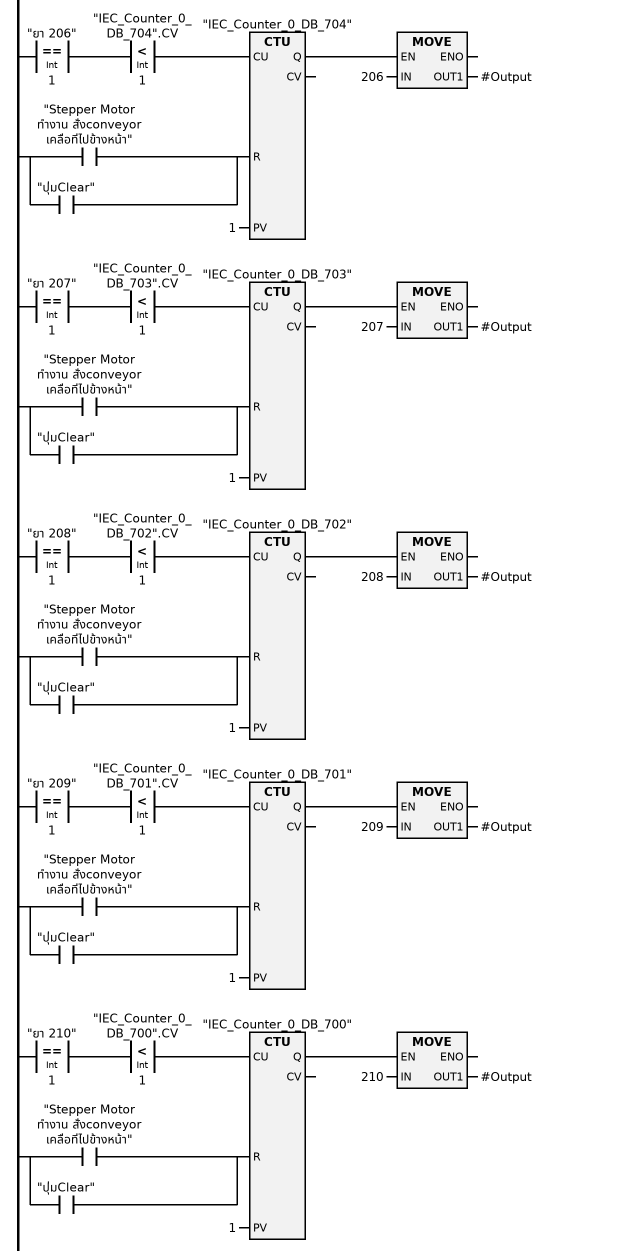
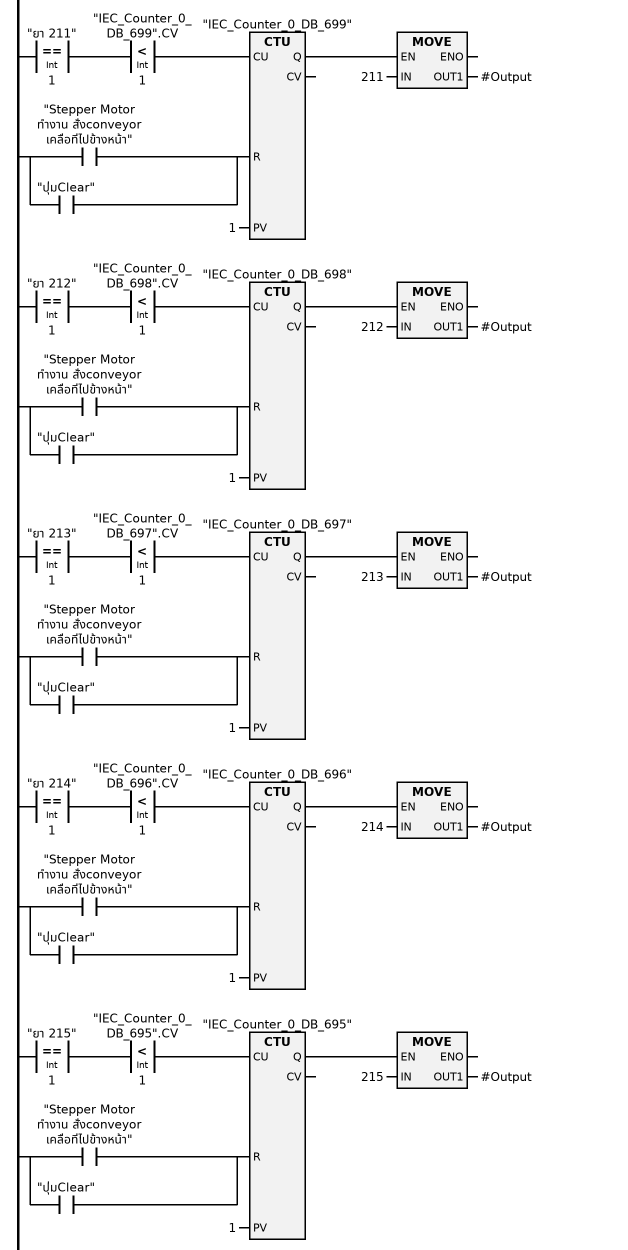
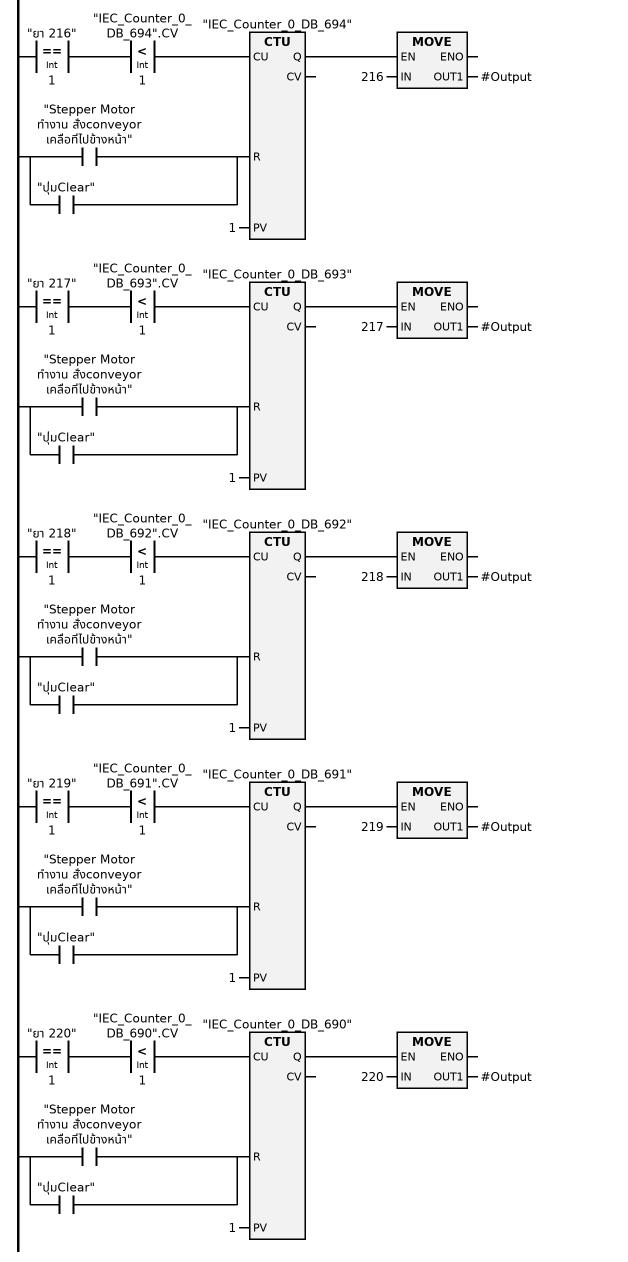
   "IEC_Counter_0_DB_709".CTU(CU := ("ยา 201" = 1) AND ("IEC_Counter_0_DB_709".CV < 1),
                           R := "Stepper Motor ทำงาน สั่งconveyor เคลื่อที่ไปข้างหน้า" OR "ปุ่มClear",
                           PV := 1);
   IF "IEC_Counter_0_DB_709".Q THEN #Output := 201; END_IF;
   "IEC_Counter_0_DB_705".CTU(CU := ("ยา 202" = 1) AND ("IEC_Counter_0_DB_705".CV < 1),
                           R := "Stepper Motor ทำงาน สั่งconveyor เคลื่อที่ไปข้างหน้า" OR "ปุ่มClear",
                           PV := 1);
   IF "IEC_Counter_0_DB_705".Q THEN #Output := 202; END_IF;
   "IEC_Counter_0_DB_708".CTU(CU := ("ยา 203" = 1) AND ("IEC_Counter_0_DB_708".CV < 1),
                           R := "Stepper Motor ทำงาน สั่งconveyor เคลื่อที่ไปข้างหน้า" OR "ปุ่มClear",
                           PV := 1);
   IF "IEC_Counter_0_DB_708".Q THEN #Output := 203; END_IF;
   "IEC_Counter_0_DB_707".CTU(CU := ("ยา 204" = 1) AND ("IEC_Counter_0_DB_707".CV < 1),
                           R := "Stepper Motor ทำงาน สั่งconveyor เคลื่อที่ไปข้างหน้า" OR "ปุ่มClear",
                           PV := 1);
   IF "IEC_Counter_0_DB_707".Q THEN #Output := 204; END_IF;
   "IEC_Counter_0_DB_706".CTU(CU := ("ยา 205" = 1) AND ("IEC_Counter_0_DB_706".CV < 1),
                           R := "Stepper Motor ทำงาน สั่งconveyor เคลื่อที่ไปข้างหน้า" OR "ปุ่มClear",
                           PV := 1);
   IF "IEC_Counter_0_DB_706".Q THEN #Output := 205; END_IF;
   "IEC_Counter_0_DB_704".CTU(CU := ("ยา 206" = 1) AND ("IEC_Counter_0_DB_704".CV < 1),
                           R := "Stepper Motor ทำงาน สั่งconveyor เคลื่อที่ไปข้างหน้า" OR "ปุ่มClear",
                           PV := 1);
   IF "IEC_Counter_0_DB_704".Q THEN #Output := 206; END_IF;
   "IEC_Counter_0_DB_703".CTU(CU := ("ยา 207" = 1) AND ("IEC_Counter_0_DB_703".CV < 1),
                           R := "Stepper Motor ทำงาน สั่งconveyor เคลื่อที่ไปข้างหน้า" OR "ปุ่มClear",
                           PV := 1);
   IF "IEC_Counter_0_DB_703".Q THEN #Output := 207; END_IF;
   "IEC_Counter_0_DB_702".CTU(CU := ("ยา 208" = 1) AND ("IEC_Counter_0_DB_702".CV < 1),
                           R := "Stepper Motor ทำงาน สั่งconveyor เคลื่อที่ไปข้างหน้า" OR "ปุ่มClear",
                           PV := 1);
   IF "IEC_Counter_0_DB_702".Q THEN #Output := 208; END_IF;
   "IEC_Counter_0_DB_701".CTU(CU := ("ยา 209" = 1) AND ("IEC_Counter_0_DB_701".CV < 1),
                           R := "Stepper Motor ทำงาน สั่งconveyor เคลื่อที่ไปข้างหน้า" OR "ปุ่มClear",
                           PV := 1);
   IF "IEC_Counter_0_DB_701".Q THEN #Output := 209; END_IF;
   "IEC_Counter_0_DB_700".CTU(CU := ("ยา 210" = 1) AND ("IEC_Counter_0_DB_700".CV < 1),
                           R := "Stepper Motor ทำงาน สั่งconveyor เคลื่อที่ไปข้างหน้า" OR "ปุ่มClear",
                           PV := 1);
   IF "IEC_Counter_0_DB_700".Q THEN #Output := 210; END_IF;
   "IEC_Counter_0_DB_699".CTU(CU := ("ยา 211" = 1) AND ("IEC_Counter_0_DB_699".CV < 1),
                           R := "Stepper Motor ทำงาน สั่งconveyor เคลื่อที่ไปข้างหน้า" OR "ปุ่มClear",
                           PV := 1);
   IF "IEC_Counter_0_DB_699".Q THEN #Output := 211; END_IF;
   "IEC_Counter_0_DB_698".CTU(CU := ("ยา 212" = 1) AND ("IEC_Counter_0_DB_698".CV < 1),
                           R := "Stepper Motor ทำงาน สั่งconveyor เคลื่อที่ไปข้างหน้า" OR "ปุ่มClear",
                           PV := 1);
   IF "IEC_Counter_0_DB_698".Q THEN #Output := 212; END_IF;
   "IEC_Counter_0_DB_697".CTU(CU := ("ยา 213" = 1) AND ("IEC_Counter_0_DB_697".CV < 1),
                           R := "Stepper Motor ทำงาน สั่งconveyor เคลื่อที่ไปข้างหน้า" OR "ปุ่มClear",
                           PV := 1);
   IF "IEC_Counter_0_DB_697".Q THEN #Output := 213; END_IF;
   "IEC_Counter_0_DB_696".CTU(CU := ("ยา 214" = 1) AND ("IEC_Counter_0_DB_696".CV < 1),
                           R := "Stepper Motor ทำงาน สั่งconveyor เคลื่อที่ไปข้างหน้า" OR "ปุ่มClear",
                           PV := 1);
   IF "IEC_Counter_0_DB_696".Q THEN #Output := 214; END_IF;
   "IEC_Counter_0_DB_695".CTU(CU := ("ยา 215" = 1) AND ("IEC_Counter_0_DB_695".CV < 1),
                           R := "Stepper Motor ทำงาน สั่งconveyor เคลื่อที่ไปข้างหน้า" OR "ปุ่มClear",
                           PV := 1);
   IF "IEC_Counter_0_DB_695".Q THEN #Output := 215; END_IF;
   "IEC_Counter_0_DB_694".CTU(CU := ("ยา 216" = 1) AND ("IEC_Counter_0_DB_694".CV < 1),
                           R := "Stepper Motor ทำงาน สั่งconveyor เคลื่อที่ไปข้างหน้า" OR "ปุ่มClear",
                           PV := 1);
   IF "IEC_Counter_0_DB_694".Q THEN #Output := 216; END_IF;
   "IEC_Counter_0_DB_693".CTU(CU := ("ยา 217" = 1) AND ("IEC_Counter_0_DB_693".CV < 1),
                           R := "Stepper Motor ทำงาน สั่งconveyor เคลื่อที่ไปข้างหน้า" OR "ปุ่มClear",
                           PV := 1);
   IF "IEC_Counter_0_DB_693".Q THEN #Output := 217; END_IF;
   "IEC_Counter_0_DB_692".CTU(CU := ("ยา 218" = 1) AND ("IEC_Counter_0_DB_692".CV < 1),
                           R := "Stepper Motor ทำงาน สั่งconveyor เคลื่อที่ไปข้างหน้า" OR "ปุ่มClear",
                           PV := 1);
   IF "IEC_Counter_0_DB_692".Q THEN #Output := 218; END_IF;
   "IEC_Counter_0_DB_691".CTU(CU := ("ยา 219" = 1) AND ("IEC_Counter_0_DB_691".CV < 1),
                           R := "Stepper Motor ทำงาน สั่งconveyor เคลื่อที่ไปข้างหน้า" OR "ปุ่มClear",
                           PV := 1);
   IF "IEC_Counter_0_DB_691".Q THEN #Output := 219; END_IF;
   "IEC_Counter_0_DB_690".CTU(CU := ("ยา 220" = 1) AND ("IEC_Counter_0_DB_690".CV < 1),
                           R := "Stepper Motor ทำงาน สั่งconveyor เคลื่อที่ไปข้างหน้า" OR "ปุ่มClear",
                           PV := 1);
   IF "IEC_Counter_0_DB_690".Q THEN #Output := 220; END_IF;
END_REGION

REGION Network 12
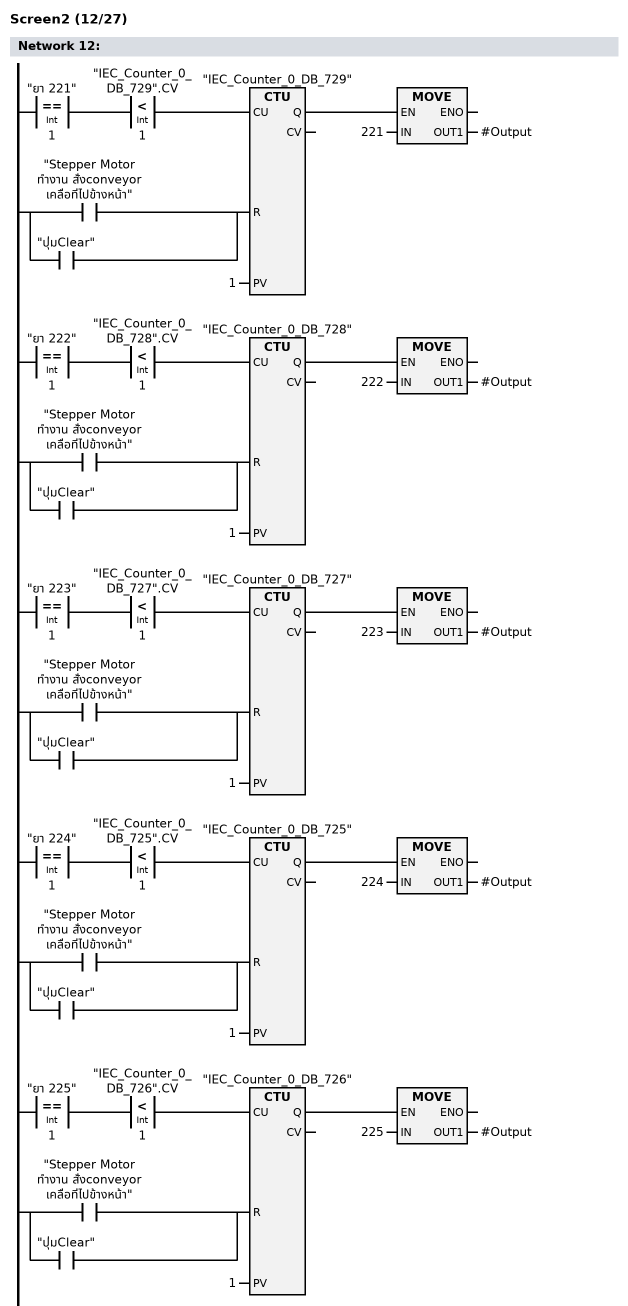
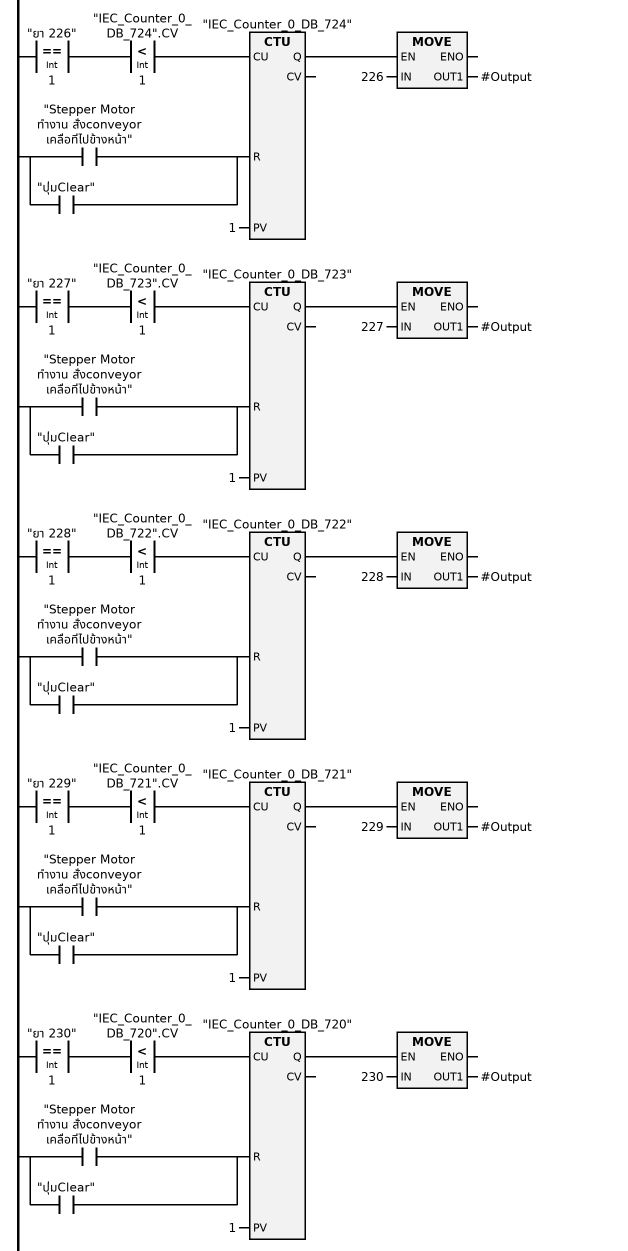
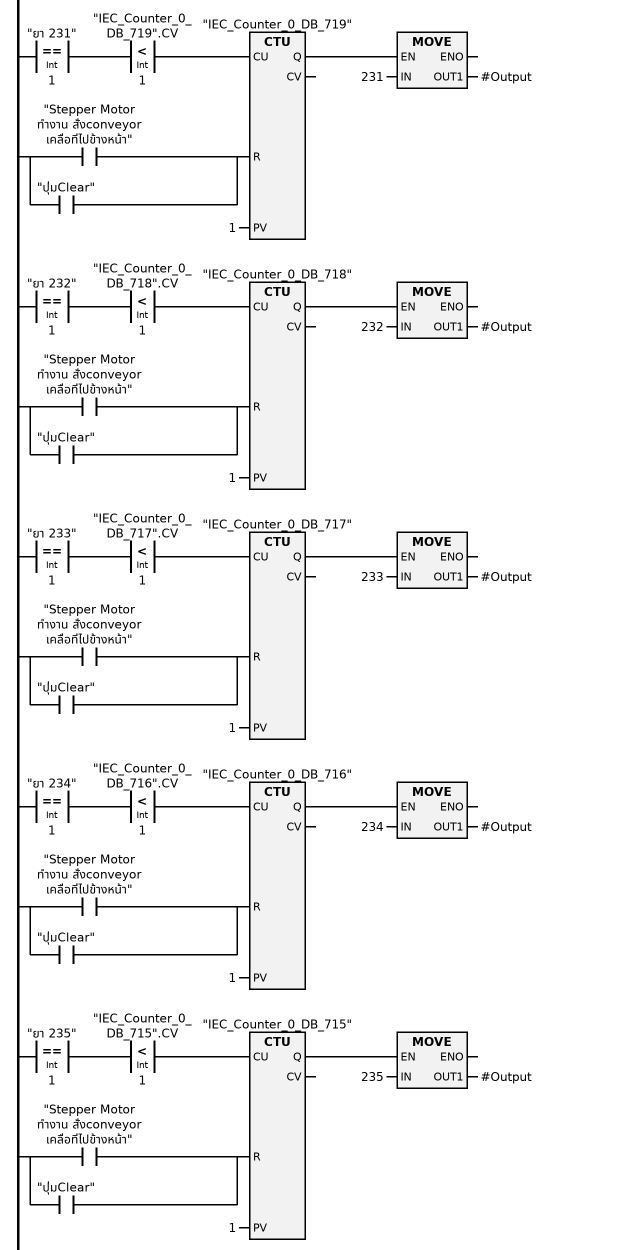
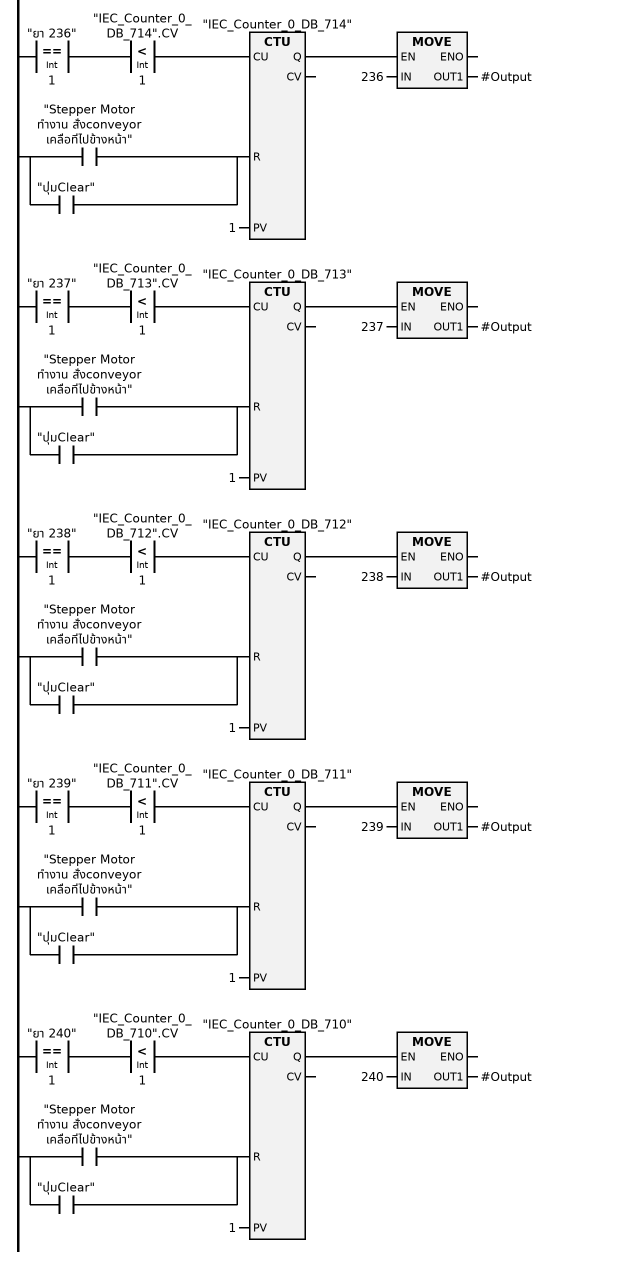
   "IEC_Counter_0_DB_729".CTU(CU := ("ยา 221" = 1) AND ("IEC_Counter_0_DB_729".CV < 1),
                           R := "Stepper Motor ทำงาน สั่งconveyor เคลื่อที่ไปข้างหน้า" OR "ปุ่มClear",
                           PV := 1);
   IF "IEC_Counter_0_DB_729".Q THEN #Output := 221; END_IF;
   "IEC_Counter_0_DB_728".CTU(CU := ("ยา 222" = 1) AND ("IEC_Counter_0_DB_728".CV < 1),
                           R := "Stepper Motor ทำงาน สั่งconveyor เคลื่อที่ไปข้างหน้า" OR "ปุ่มClear",
                           PV := 1);
   IF "IEC_Counter_0_DB_728".Q THEN #Output := 222; END_IF;
   "IEC_Counter_0_DB_727".CTU(CU := ("ยา 223" = 1) AND ("IEC_Counter_0_DB_727".CV < 1),
                           R := "Stepper Motor ทำงาน สั่งconveyor เคลื่อที่ไปข้างหน้า" OR "ปุ่มClear",
                           PV := 1);
   IF "IEC_Counter_0_DB_727".Q THEN #Output := 223; END_IF;
   "IEC_Counter_0_DB_725".CTU(CU := ("ยา 224" = 1) AND ("IEC_Counter_0_DB_725".CV < 1),
                           R := "Stepper Motor ทำงาน สั่งconveyor เคลื่อที่ไปข้างหน้า" OR "ปุ่มClear",
                           PV := 1);
   IF "IEC_Counter_0_DB_725".Q THEN #Output := 224; END_IF;
   "IEC_Counter_0_DB_726".CTU(CU := ("ยา 225" = 1) AND ("IEC_Counter_0_DB_726".CV < 1),
                           R := "Stepper Motor ทำงาน สั่งconveyor เคลื่อที่ไปข้างหน้า" OR "ปุ่มClear",
                           PV := 1);
   IF "IEC_Counter_0_DB_726".Q THEN #Output := 225; END_IF;
   "IEC_Counter_0_DB_724".CTU(CU := ("ยา 226" = 1) AND ("IEC_Counter_0_DB_724".CV < 1),
                           R := "Stepper Motor ทำงาน สั่งconveyor เคลื่อที่ไปข้างหน้า" OR "ปุ่มClear",
                           PV := 1);
   IF "IEC_Counter_0_DB_724".Q THEN #Output := 226; END_IF;
   "IEC_Counter_0_DB_723".CTU(CU := ("ยา 227" = 1) AND ("IEC_Counter_0_DB_723".CV < 1),
                           R := "Stepper Motor ทำงาน สั่งconveyor เคลื่อที่ไปข้างหน้า" OR "ปุ่มClear",
                           PV := 1);
   IF "IEC_Counter_0_DB_723".Q THEN #Output := 227; END_IF;
   "IEC_Counter_0_DB_722".CTU(CU := ("ยา 228" = 1) AND ("IEC_Counter_0_DB_722".CV < 1),
                           R := "Stepper Motor ทำงาน สั่งconveyor เคลื่อที่ไปข้างหน้า" OR "ปุ่มClear",
                           PV := 1);
   IF "IEC_Counter_0_DB_722".Q THEN #Output := 228; END_IF;
   "IEC_Counter_0_DB_721".CTU(CU := ("ยา 229" = 1) AND ("IEC_Counter_0_DB_721".CV < 1),
                           R := "Stepper Motor ทำงาน สั่งconveyor เคลื่อที่ไปข้างหน้า" OR "ปุ่มClear",
                           PV := 1);
   IF "IEC_Counter_0_DB_721".Q THEN #Output := 229; END_IF;
   "IEC_Counter_0_DB_720".CTU(CU := ("ยา 230" = 1) AND ("IEC_Counter_0_DB_720".CV < 1),
                           R := "Stepper Motor ทำงาน สั่งconveyor เคลื่อที่ไปข้างหน้า" OR "ปุ่มClear",
                           PV := 1);
   IF "IEC_Counter_0_DB_720".Q THEN #Output := 230; END_IF;
   "IEC_Counter_0_DB_719".CTU(CU := ("ยา 231" = 1) AND ("IEC_Counter_0_DB_719".CV < 1),
                           R := "Stepper Motor ทำงาน สั่งconveyor เคลื่อที่ไปข้างหน้า" OR "ปุ่มClear",
                           PV := 1);
   IF "IEC_Counter_0_DB_719".Q THEN #Output := 231; END_IF;
   "IEC_Counter_0_DB_718".CTU(CU := ("ยา 232" = 1) AND ("IEC_Counter_0_DB_718".CV < 1),
                           R := "Stepper Motor ทำงาน สั่งconveyor เคลื่อที่ไปข้างหน้า" OR "ปุ่มClear",
                           PV := 1);
   IF "IEC_Counter_0_DB_718".Q THEN #Output := 232; END_IF;
   "IEC_Counter_0_DB_717".CTU(CU := ("ยา 233" = 1) AND ("IEC_Counter_0_DB_717".CV < 1),
                           R := "Stepper Motor ทำงาน สั่งconveyor เคลื่อที่ไปข้างหน้า" OR "ปุ่มClear",
                           PV := 1);
   IF "IEC_Counter_0_DB_717".Q THEN #Output := 233; END_IF;
   "IEC_Counter_0_DB_716".CTU(CU := ("ยา 234" = 1) AND ("IEC_Counter_0_DB_716".CV < 1),
                           R := "Stepper Motor ทำงาน สั่งconveyor เคลื่อที่ไปข้างหน้า" OR "ปุ่มClear",
                           PV := 1);
   IF "IEC_Counter_0_DB_716".Q THEN #Output := 234; END_IF;
   "IEC_Counter_0_DB_715".CTU(CU := ("ยา 235" = 1) AND ("IEC_Counter_0_DB_715".CV < 1),
                           R := "Stepper Motor ทำงาน สั่งconveyor เคลื่อที่ไปข้างหน้า" OR "ปุ่มClear",
                           PV := 1);
   IF "IEC_Counter_0_DB_715".Q THEN #Output := 235; END_IF;
   "IEC_Counter_0_DB_714".CTU(CU := ("ยา 236" = 1) AND ("IEC_Counter_0_DB_714".CV < 1),
                           R := "Stepper Motor ทำงาน สั่งconveyor เคลื่อที่ไปข้างหน้า" OR "ปุ่มClear",
                           PV := 1);
   IF "IEC_Counter_0_DB_714".Q THEN #Output := 236; END_IF;
   "IEC_Counter_0_DB_713".CTU(CU := ("ยา 237" = 1) AND ("IEC_Counter_0_DB_713".CV < 1),
                           R := "Stepper Motor ทำงาน สั่งconveyor เคลื่อที่ไปข้างหน้า" OR "ปุ่มClear",
                           PV := 1);
   IF "IEC_Counter_0_DB_713".Q THEN #Output := 237; END_IF;
   "IEC_Counter_0_DB_712".CTU(CU := ("ยา 238" = 1) AND ("IEC_Counter_0_DB_712".CV < 1),
                           R := "Stepper Motor ทำงาน สั่งconveyor เคลื่อที่ไปข้างหน้า" OR "ปุ่มClear",
                           PV := 1);
   IF "IEC_Counter_0_DB_712".Q THEN #Output := 238; END_IF;
   "IEC_Counter_0_DB_711".CTU(CU := ("ยา 239" = 1) AND ("IEC_Counter_0_DB_711".CV < 1),
                           R := "Stepper Motor ทำงาน สั่งconveyor เคลื่อที่ไปข้างหน้า" OR "ปุ่มClear",
                           PV := 1);
   IF "IEC_Counter_0_DB_711".Q THEN #Output := 239; END_IF;
   "IEC_Counter_0_DB_710".CTU(CU := ("ยา 240" = 1) AND ("IEC_Counter_0_DB_710".CV < 1),
                           R := "Stepper Motor ทำงาน สั่งconveyor เคลื่อที่ไปข้างหน้า" OR "ปุ่มClear",
                           PV := 1);
   IF "IEC_Counter_0_DB_710".Q THEN #Output := 240; END_IF;
END_REGION

REGION Network 13
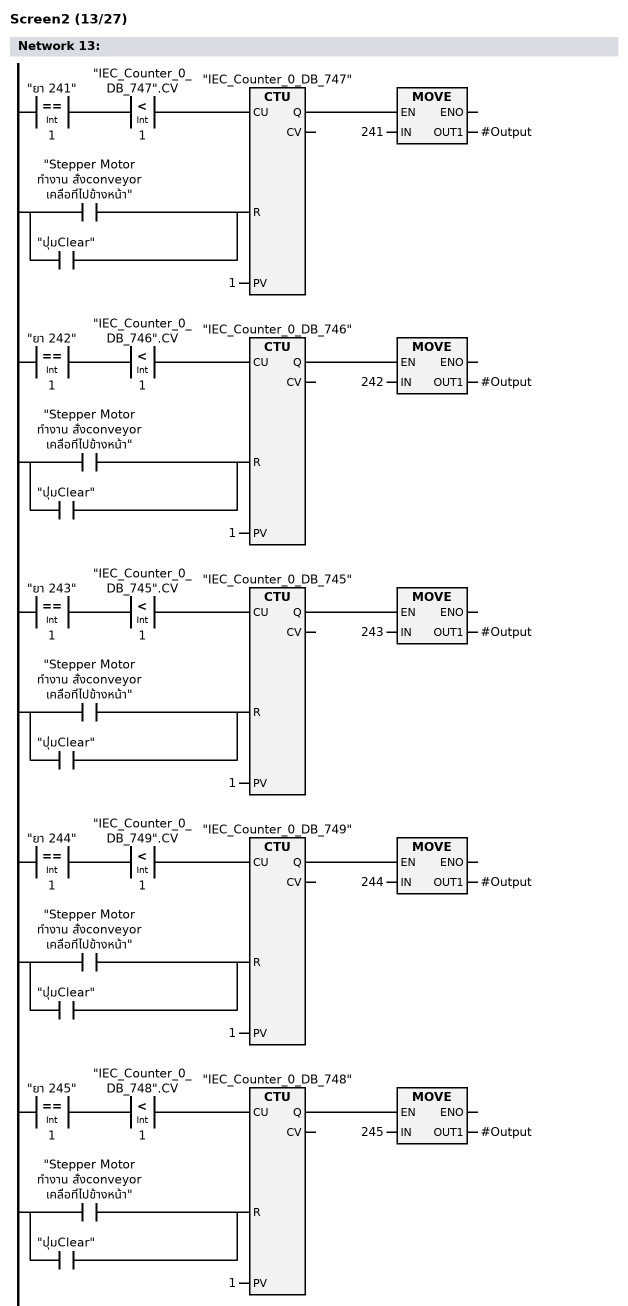
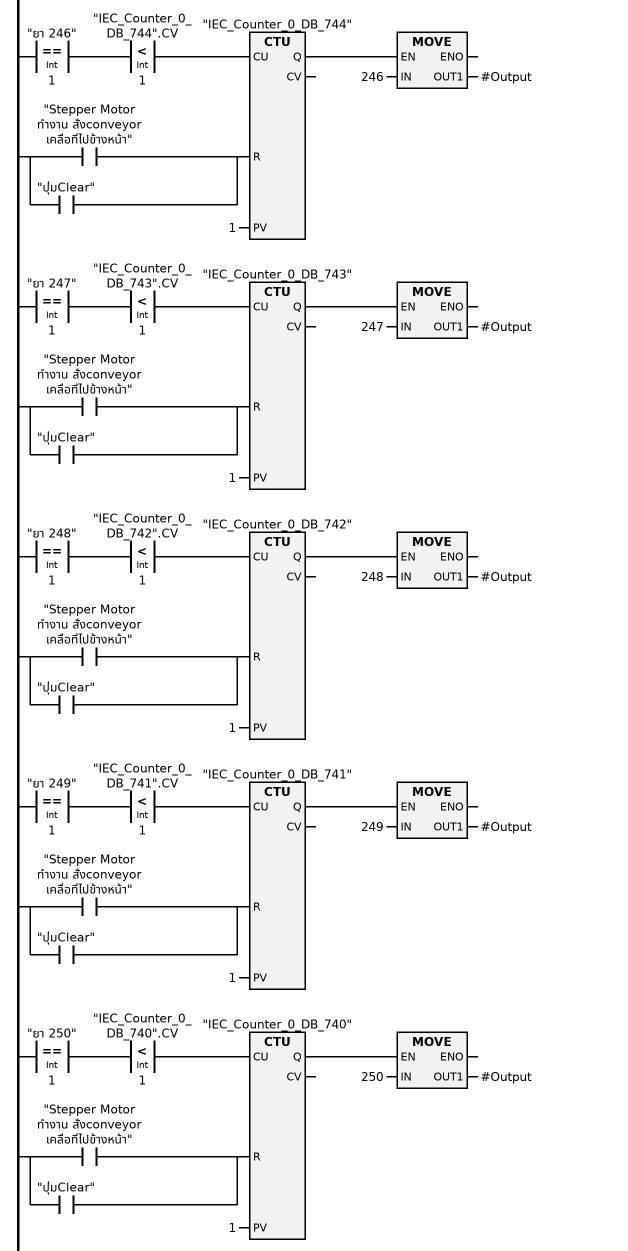
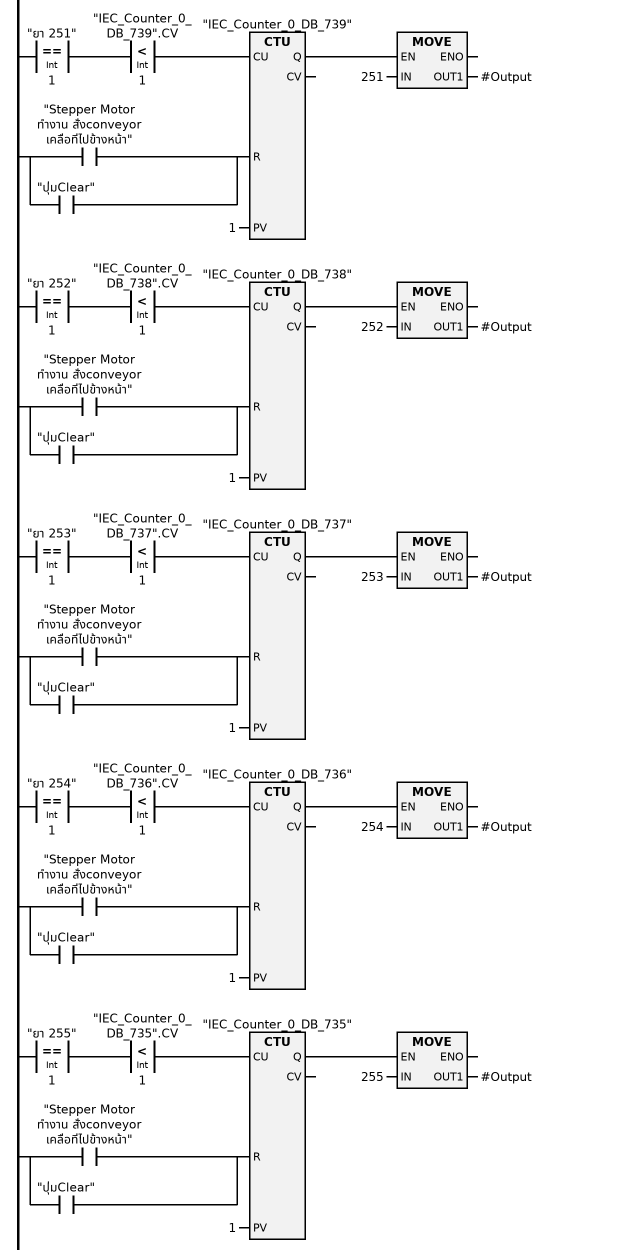
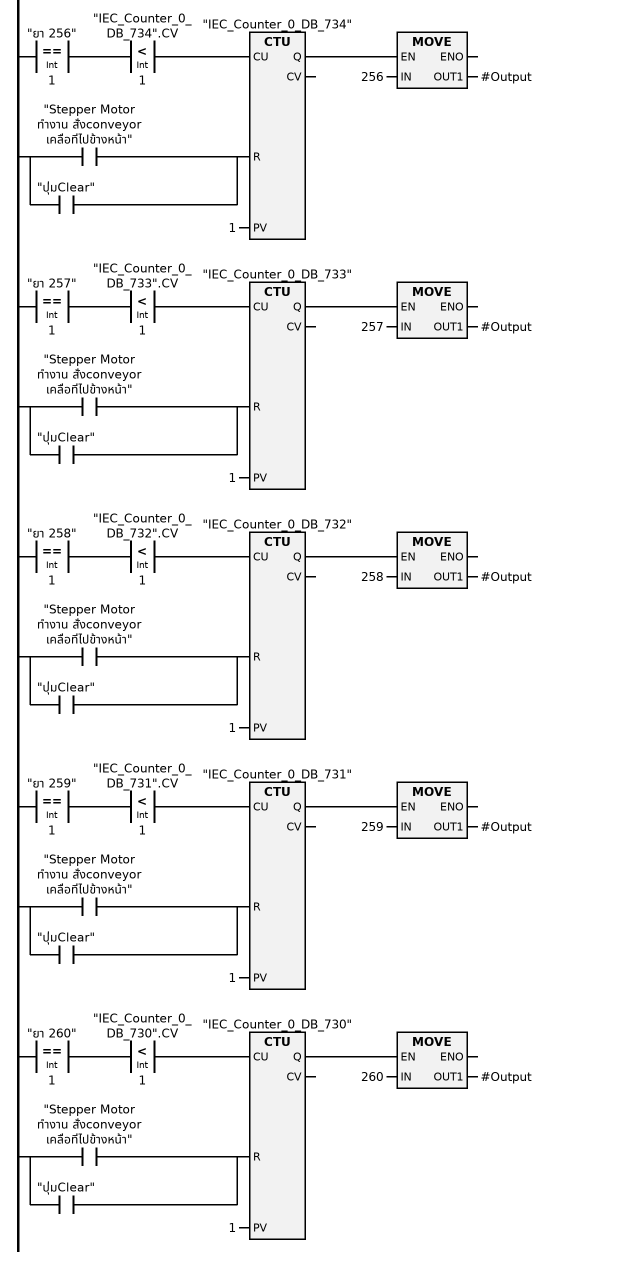
   "IEC_Counter_0_DB_747".CTU(CU := ("ยา 241" = 1) AND ("IEC_Counter_0_DB_747".CV < 1),
                           R := "Stepper Motor ทำงาน สั่งconveyor เคลื่อที่ไปข้างหน้า" OR "ปุ่มClear",
                           PV := 1);
   IF "IEC_Counter_0_DB_747".Q THEN #Output := 241; END_IF;
   "IEC_Counter_0_DB_746".CTU(CU := ("ยา 242" = 1) AND ("IEC_Counter_0_DB_746".CV < 1),
                           R := "Stepper Motor ทำงาน สั่งconveyor เคลื่อที่ไปข้างหน้า" OR "ปุ่มClear",
                           PV := 1);
   IF "IEC_Counter_0_DB_746".Q THEN #Output := 242; END_IF;
   "IEC_Counter_0_DB_745".CTU(CU := ("ยา 243" = 1) AND ("IEC_Counter_0_DB_745".CV < 1),
                           R := "Stepper Motor ทำงาน สั่งconveyor เคลื่อที่ไปข้างหน้า" OR "ปุ่มClear",
                           PV := 1);
   IF "IEC_Counter_0_DB_745".Q THEN #Output := 243; END_IF;
   "IEC_Counter_0_DB_749".CTU(CU := ("ยา 244" = 1) AND ("IEC_Counter_0_DB_749".CV < 1),
                           R := "Stepper Motor ทำงาน สั่งconveyor เคลื่อที่ไปข้างหน้า" OR "ปุ่มClear",
                           PV := 1);
   IF "IEC_Counter_0_DB_749".Q THEN #Output := 244; END_IF;
   "IEC_Counter_0_DB_748".CTU(CU := ("ยา 245" = 1) AND ("IEC_Counter_0_DB_748".CV < 1),
                           R := "Stepper Motor ทำงาน สั่งconveyor เคลื่อที่ไปข้างหน้า" OR "ปุ่มClear",
                           PV := 1);
   IF "IEC_Counter_0_DB_748".Q THEN #Output := 245; END_IF;
   "IEC_Counter_0_DB_744".CTU(CU := ("ยา 246" = 1) AND ("IEC_Counter_0_DB_744".CV < 1),
                           R := "Stepper Motor ทำงาน สั่งconveyor เคลื่อที่ไปข้างหน้า" OR "ปุ่มClear",
                           PV := 1);
   IF "IEC_Counter_0_DB_744".Q THEN #Output := 246; END_IF;
   "IEC_Counter_0_DB_743".CTU(CU := ("ยา 247" = 1) AND ("IEC_Counter_0_DB_743".CV < 1),
                           R := "Stepper Motor ทำงาน สั่งconveyor เคลื่อที่ไปข้างหน้า" OR "ปุ่มClear",
                           PV := 1);
   IF "IEC_Counter_0_DB_743".Q THEN #Output := 247; END_IF;
   "IEC_Counter_0_DB_742".CTU(CU := ("ยา 248" = 1) AND ("IEC_Counter_0_DB_742".CV < 1),
                           R := "Stepper Motor ทำงาน สั่งconveyor เคลื่อที่ไปข้างหน้า" OR "ปุ่มClear",
                           PV := 1);
   IF "IEC_Counter_0_DB_742".Q THEN #Output := 248; END_IF;
   "IEC_Counter_0_DB_741".CTU(CU := ("ยา 249" = 1) AND ("IEC_Counter_0_DB_741".CV < 1),
                           R := "Stepper Motor ทำงาน สั่งconveyor เคลื่อที่ไปข้างหน้า" OR "ปุ่มClear",
                           PV := 1);
   IF "IEC_Counter_0_DB_741".Q THEN #Output := 249; END_IF;
   "IEC_Counter_0_DB_740".CTU(CU := ("ยา 250" = 1) AND ("IEC_Counter_0_DB_740".CV < 1),
                           R := "Stepper Motor ทำงาน สั่งconveyor เคลื่อที่ไปข้างหน้า" OR "ปุ่มClear",
                           PV := 1);
   IF "IEC_Counter_0_DB_740".Q THEN #Output := 250; END_IF;
   "IEC_Counter_0_DB_739".CTU(CU := ("ยา 251" = 1) AND ("IEC_Counter_0_DB_739".CV < 1),
                           R := "Stepper Motor ทำงาน สั่งconveyor เคลื่อที่ไปข้างหน้า" OR "ปุ่มClear",
                           PV := 1);
   IF "IEC_Counter_0_DB_739".Q THEN #Output := 251; END_IF;
   "IEC_Counter_0_DB_738".CTU(CU := ("ยา 252" = 1) AND ("IEC_Counter_0_DB_738".CV < 1),
                           R := "Stepper Motor ทำงาน สั่งconveyor เคลื่อที่ไปข้างหน้า" OR "ปุ่มClear",
                           PV := 1);
   IF "IEC_Counter_0_DB_738".Q THEN #Output := 252; END_IF;
   "IEC_Counter_0_DB_737".CTU(CU := ("ยา 253" = 1) AND ("IEC_Counter_0_DB_737".CV < 1),
                           R := "Stepper Motor ทำงาน สั่งconveyor เคลื่อที่ไปข้างหน้า" OR "ปุ่มClear",
                           PV := 1);
   IF "IEC_Counter_0_DB_737".Q THEN #Output := 253; END_IF;
   "IEC_Counter_0_DB_736".CTU(CU := ("ยา 254" = 1) AND ("IEC_Counter_0_DB_736".CV < 1),
                           R := "Stepper Motor ทำงาน สั่งconveyor เคลื่อที่ไปข้างหน้า" OR "ปุ่มClear",
                           PV := 1);
   IF "IEC_Counter_0_DB_736".Q THEN #Output := 254; END_IF;
   "IEC_Counter_0_DB_735".CTU(CU := ("ยา 255" = 1) AND ("IEC_Counter_0_DB_735".CV < 1),
                           R := "Stepper Motor ทำงาน สั่งconveyor เคลื่อที่ไปข้างหน้า" OR "ปุ่มClear",
                           PV := 1);
   IF "IEC_Counter_0_DB_735".Q THEN #Output := 255; END_IF;
   "IEC_Counter_0_DB_734".CTU(CU := ("ยา 256" = 1) AND ("IEC_Counter_0_DB_734".CV < 1),
                           R := "Stepper Motor ทำงาน สั่งconveyor เคลื่อที่ไปข้างหน้า" OR "ปุ่มClear",
                           PV := 1);
   IF "IEC_Counter_0_DB_734".Q THEN #Output := 256; END_IF;
   "IEC_Counter_0_DB_733".CTU(CU := ("ยา 257" = 1) AND ("IEC_Counter_0_DB_733".CV < 1),
                           R := "Stepper Motor ทำงาน สั่งconveyor เคลื่อที่ไปข้างหน้า" OR "ปุ่มClear",
                           PV := 1);
   IF "IEC_Counter_0_DB_733".Q THEN #Output := 257; END_IF;
   "IEC_Counter_0_DB_732".CTU(CU := ("ยา 258" = 1) AND ("IEC_Counter_0_DB_732".CV < 1),
                           R := "Stepper Motor ทำงาน สั่งconveyor เคลื่อที่ไปข้างหน้า" OR "ปุ่มClear",
                           PV := 1);
   IF "IEC_Counter_0_DB_732".Q THEN #Output := 258; END_IF;
   "IEC_Counter_0_DB_731".CTU(CU := ("ยา 259" = 1) AND ("IEC_Counter_0_DB_731".CV < 1),
                           R := "Stepper Motor ทำงาน สั่งconveyor เคลื่อที่ไปข้างหน้า" OR "ปุ่มClear",
                           PV := 1);
   IF "IEC_Counter_0_DB_731".Q THEN #Output := 259; END_IF;
   "IEC_Counter_0_DB_730".CTU(CU := ("ยา 260" = 1) AND ("IEC_Counter_0_DB_730".CV < 1),
                           R := "Stepper Motor ทำงาน สั่งconveyor เคลื่อที่ไปข้างหน้า" OR "ปุ่มClear",
                           PV := 1);
   IF "IEC_Counter_0_DB_730".Q THEN #Output := 260; END_IF;
END_REGION

REGION Network 14
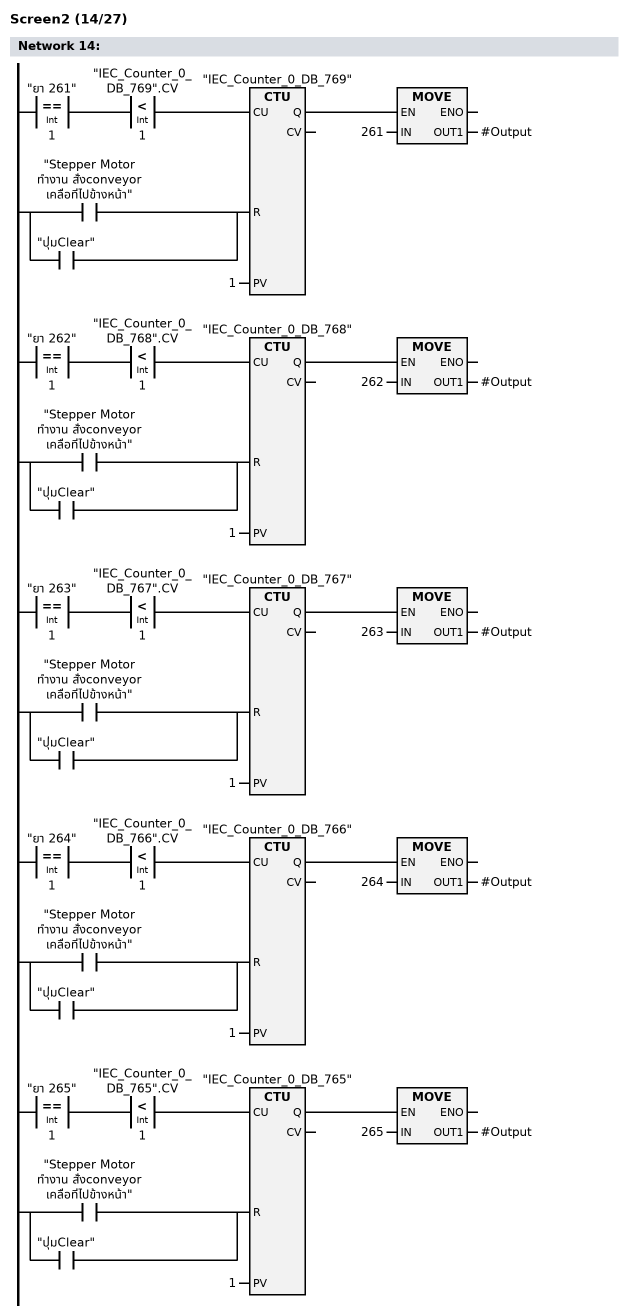
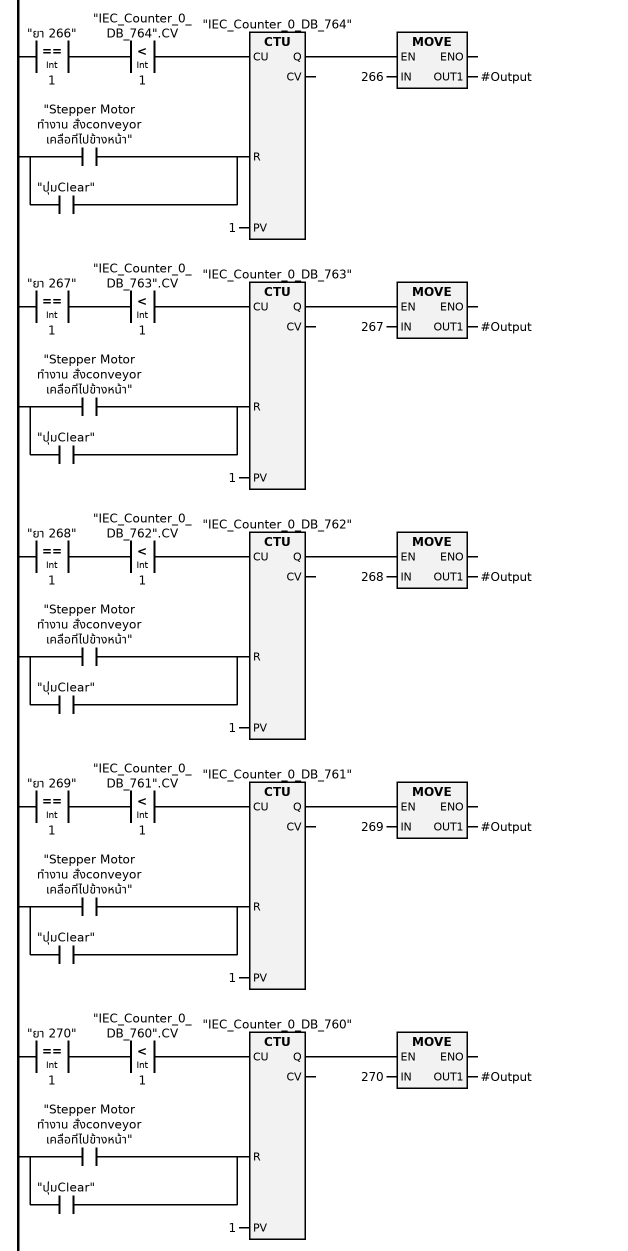
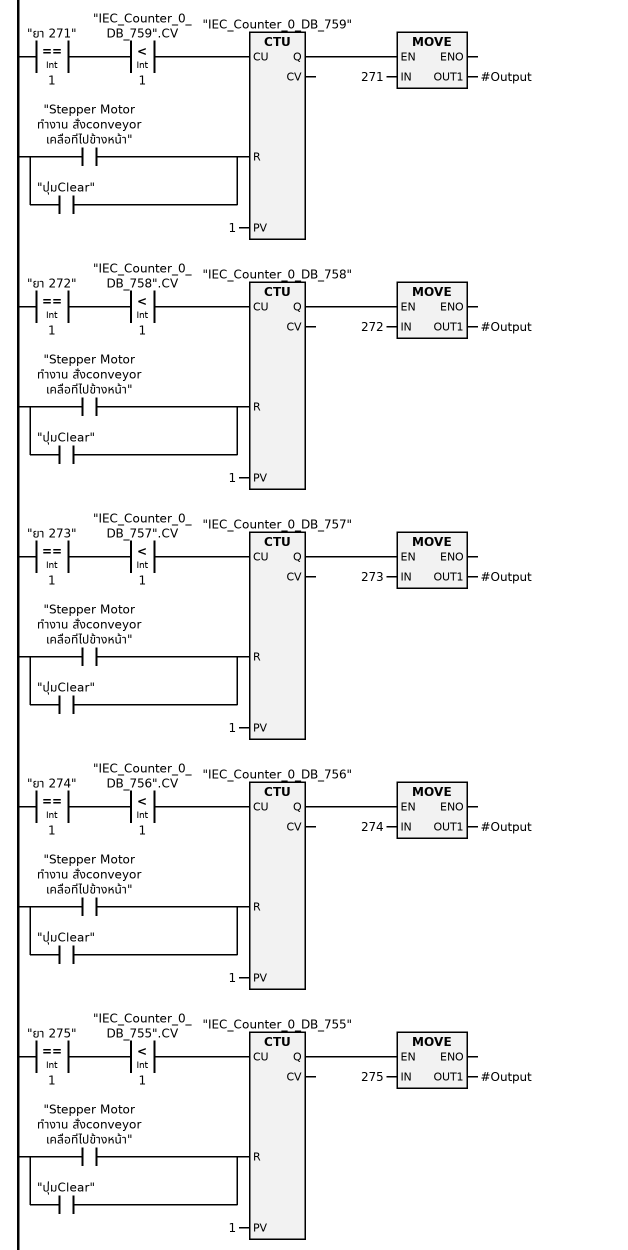
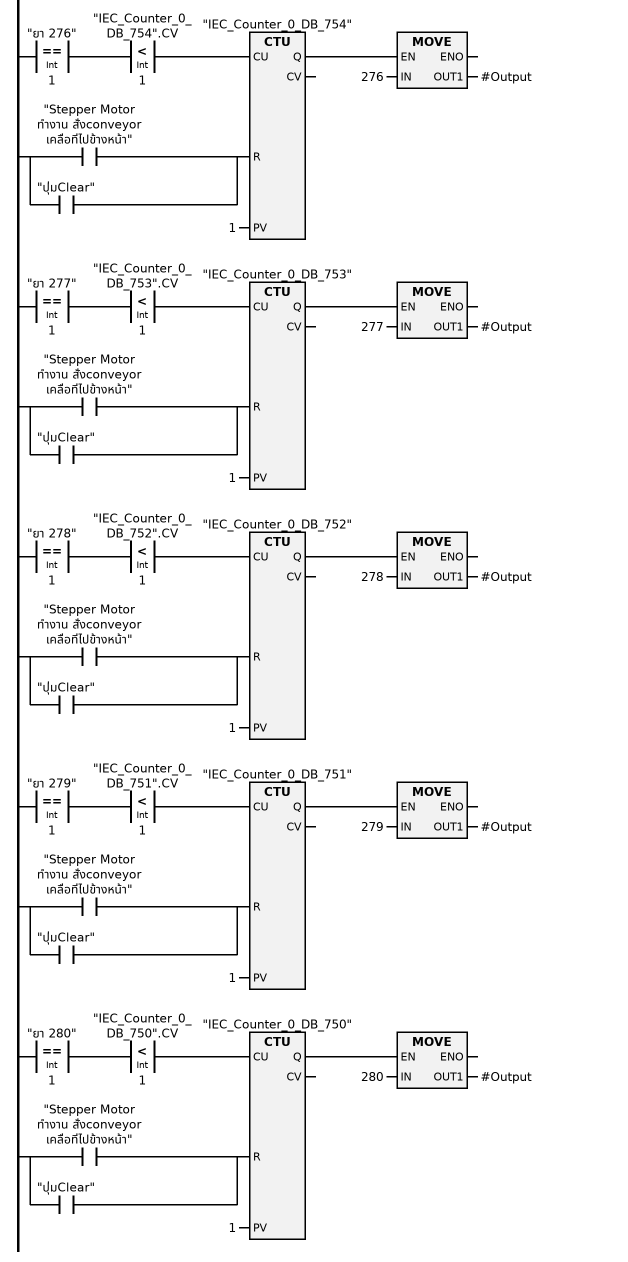
   "IEC_Counter_0_DB_769".CTU(CU := ("ยา 261" = 1) AND ("IEC_Counter_0_DB_769".CV < 1),
                           R := "Stepper Motor ทำงาน สั่งconveyor เคลื่อที่ไปข้างหน้า" OR "ปุ่มClear",
                           PV := 1);
   IF "IEC_Counter_0_DB_769".Q THEN #Output := 261; END_IF;
   "IEC_Counter_0_DB_768".CTU(CU := ("ยา 262" = 1) AND ("IEC_Counter_0_DB_768".CV < 1),
                           R := "Stepper Motor ทำงาน สั่งconveyor เคลื่อที่ไปข้างหน้า" OR "ปุ่มClear",
                           PV := 1);
   IF "IEC_Counter_0_DB_768".Q THEN #Output := 262; END_IF;
   "IEC_Counter_0_DB_767".CTU(CU := ("ยา 263" = 1) AND ("IEC_Counter_0_DB_767".CV < 1),
                           R := "Stepper Motor ทำงาน สั่งconveyor เคลื่อที่ไปข้างหน้า" OR "ปุ่มClear",
                           PV := 1);
   IF "IEC_Counter_0_DB_767".Q THEN #Output := 263; END_IF;
   "IEC_Counter_0_DB_766".CTU(CU := ("ยา 264" = 1) AND ("IEC_Counter_0_DB_766".CV < 1),
                           R := "Stepper Motor ทำงาน สั่งconveyor เคลื่อที่ไปข้างหน้า" OR "ปุ่มClear",
                           PV := 1);
   IF "IEC_Counter_0_DB_766".Q THEN #Output := 264; END_IF;
   "IEC_Counter_0_DB_765".CTU(CU := ("ยา 265" = 1) AND ("IEC_Counter_0_DB_765".CV < 1),
                           R := "Stepper Motor ทำงาน สั่งconveyor เคลื่อที่ไปข้างหน้า" OR "ปุ่มClear",
                           PV := 1);
   IF "IEC_Counter_0_DB_765".Q THEN #Output := 265; END_IF;
   "IEC_Counter_0_DB_764".CTU(CU := ("ยา 266" = 1) AND ("IEC_Counter_0_DB_764".CV < 1),
                           R := "Stepper Motor ทำงาน สั่งconveyor เคลื่อที่ไปข้างหน้า" OR "ปุ่มClear",
                           PV := 1);
   IF "IEC_Counter_0_DB_764".Q THEN #Output := 266; END_IF;
   "IEC_Counter_0_DB_763".CTU(CU := ("ยา 267" = 1) AND ("IEC_Counter_0_DB_763".CV < 1),
                           R := "Stepper Motor ทำงาน สั่งconveyor เคลื่อที่ไปข้างหน้า" OR "ปุ่มClear",
                           PV := 1);
   IF "IEC_Counter_0_DB_763".Q THEN #Output := 267; END_IF;
   "IEC_Counter_0_DB_762".CTU(CU := ("ยา 268" = 1) AND ("IEC_Counter_0_DB_762".CV < 1),
                           R := "Stepper Motor ทำงาน สั่งconveyor เคลื่อที่ไปข้างหน้า" OR "ปุ่มClear",
                           PV := 1);
   IF "IEC_Counter_0_DB_762".Q THEN #Output := 268; END_IF;
   "IEC_Counter_0_DB_761".CTU(CU := ("ยา 269" = 1) AND ("IEC_Counter_0_DB_761".CV < 1),
                           R := "Stepper Motor ทำงาน สั่งconveyor เคลื่อที่ไปข้างหน้า" OR "ปุ่มClear",
                           PV := 1);
   IF "IEC_Counter_0_DB_761".Q THEN #Output := 269; END_IF;
   "IEC_Counter_0_DB_760".CTU(CU := ("ยา 270" = 1) AND ("IEC_Counter_0_DB_760".CV < 1),
                           R := "Stepper Motor ทำงาน สั่งconveyor เคลื่อที่ไปข้างหน้า" OR "ปุ่มClear",
                           PV := 1);
   IF "IEC_Counter_0_DB_760".Q THEN #Output := 270; END_IF;
   "IEC_Counter_0_DB_759".CTU(CU := ("ยา 271" = 1) AND ("IEC_Counter_0_DB_759".CV < 1),
                           R := "Stepper Motor ทำงาน สั่งconveyor เคลื่อที่ไปข้างหน้า" OR "ปุ่มClear",
                           PV := 1);
   IF "IEC_Counter_0_DB_759".Q THEN #Output := 271; END_IF;
   "IEC_Counter_0_DB_758".CTU(CU := ("ยา 272" = 1) AND ("IEC_Counter_0_DB_758".CV < 1),
                           R := "Stepper Motor ทำงาน สั่งconveyor เคลื่อที่ไปข้างหน้า" OR "ปุ่มClear",
                           PV := 1);
   IF "IEC_Counter_0_DB_758".Q THEN #Output := 272; END_IF;
   "IEC_Counter_0_DB_757".CTU(CU := ("ยา 273" = 1) AND ("IEC_Counter_0_DB_757".CV < 1),
                           R := "Stepper Motor ทำงาน สั่งconveyor เคลื่อที่ไปข้างหน้า" OR "ปุ่มClear",
                           PV := 1);
   IF "IEC_Counter_0_DB_757".Q THEN #Output := 273; END_IF;
   "IEC_Counter_0_DB_756".CTU(CU := ("ยา 274" = 1) AND ("IEC_Counter_0_DB_756".CV < 1),
                           R := "Stepper Motor ทำงาน สั่งconveyor เคลื่อที่ไปข้างหน้า" OR "ปุ่มClear",
                           PV := 1);
   IF "IEC_Counter_0_DB_756".Q THEN #Output := 274; END_IF;
   "IEC_Counter_0_DB_755".CTU(CU := ("ยา 275" = 1) AND ("IEC_Counter_0_DB_755".CV < 1),
                           R := "Stepper Motor ทำงาน สั่งconveyor เคลื่อที่ไปข้างหน้า" OR "ปุ่มClear",
                           PV := 1);
   IF "IEC_Counter_0_DB_755".Q THEN #Output := 275; END_IF;
   "IEC_Counter_0_DB_754".CTU(CU := ("ยา 276" = 1) AND ("IEC_Counter_0_DB_754".CV < 1),
                           R := "Stepper Motor ทำงาน สั่งconveyor เคลื่อที่ไปข้างหน้า" OR "ปุ่มClear",
                           PV := 1);
   IF "IEC_Counter_0_DB_754".Q THEN #Output := 276; END_IF;
   "IEC_Counter_0_DB_753".CTU(CU := ("ยา 277" = 1) AND ("IEC_Counter_0_DB_753".CV < 1),
                           R := "Stepper Motor ทำงาน สั่งconveyor เคลื่อที่ไปข้างหน้า" OR "ปุ่มClear",
                           PV := 1);
   IF "IEC_Counter_0_DB_753".Q THEN #Output := 277; END_IF;
   "IEC_Counter_0_DB_752".CTU(CU := ("ยา 278" = 1) AND ("IEC_Counter_0_DB_752".CV < 1),
                           R := "Stepper Motor ทำงาน สั่งconveyor เคลื่อที่ไปข้างหน้า" OR "ปุ่มClear",
                           PV := 1);
   IF "IEC_Counter_0_DB_752".Q THEN #Output := 278; END_IF;
   "IEC_Counter_0_DB_751".CTU(CU := ("ยา 279" = 1) AND ("IEC_Counter_0_DB_751".CV < 1),
                           R := "Stepper Motor ทำงาน สั่งconveyor เคลื่อที่ไปข้างหน้า" OR "ปุ่มClear",
                           PV := 1);
   IF "IEC_Counter_0_DB_751".Q THEN #Output := 279; END_IF;
   "IEC_Counter_0_DB_750".CTU(CU := ("ยา 280" = 1) AND ("IEC_Counter_0_DB_750".CV < 1),
                           R := "Stepper Motor ทำงาน สั่งconveyor เคลื่อที่ไปข้างหน้า" OR "ปุ่มClear",
                           PV := 1);
   IF "IEC_Counter_0_DB_750".Q THEN #Output := 280; END_IF;
END_REGION

REGION Network 15
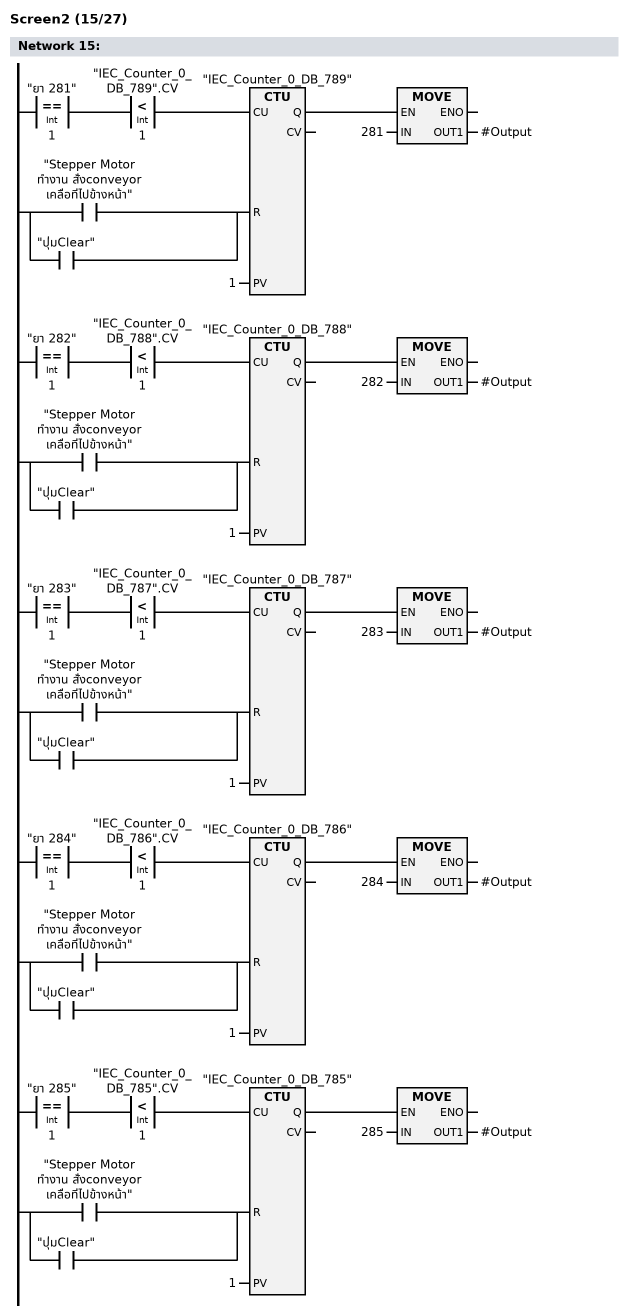
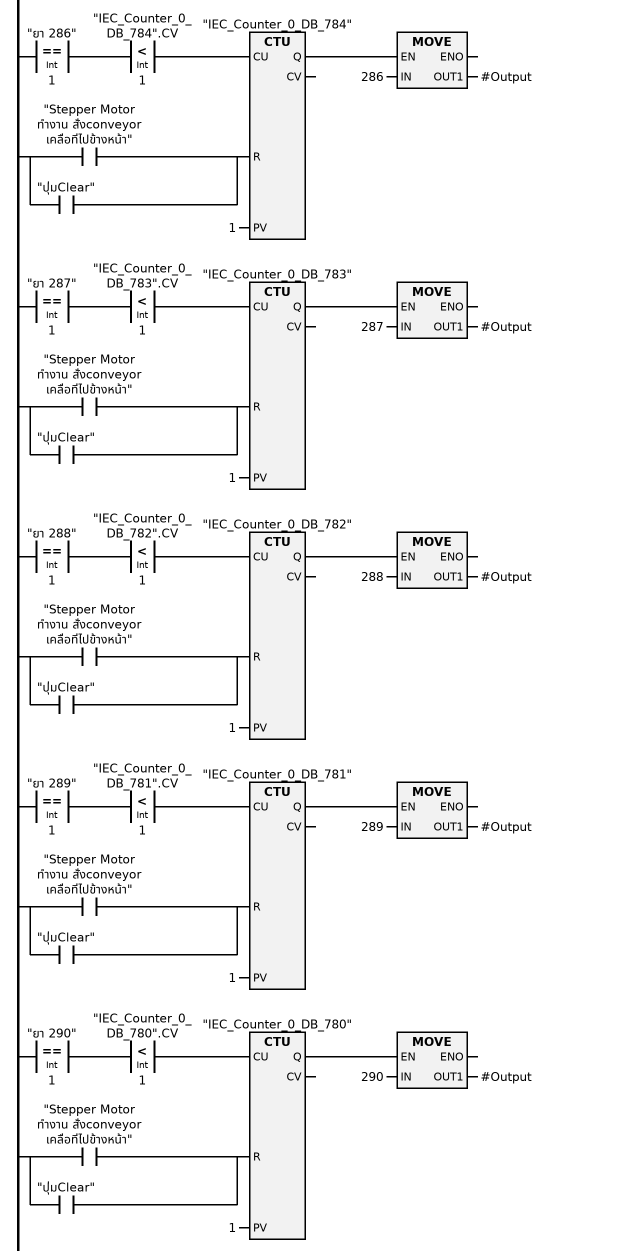
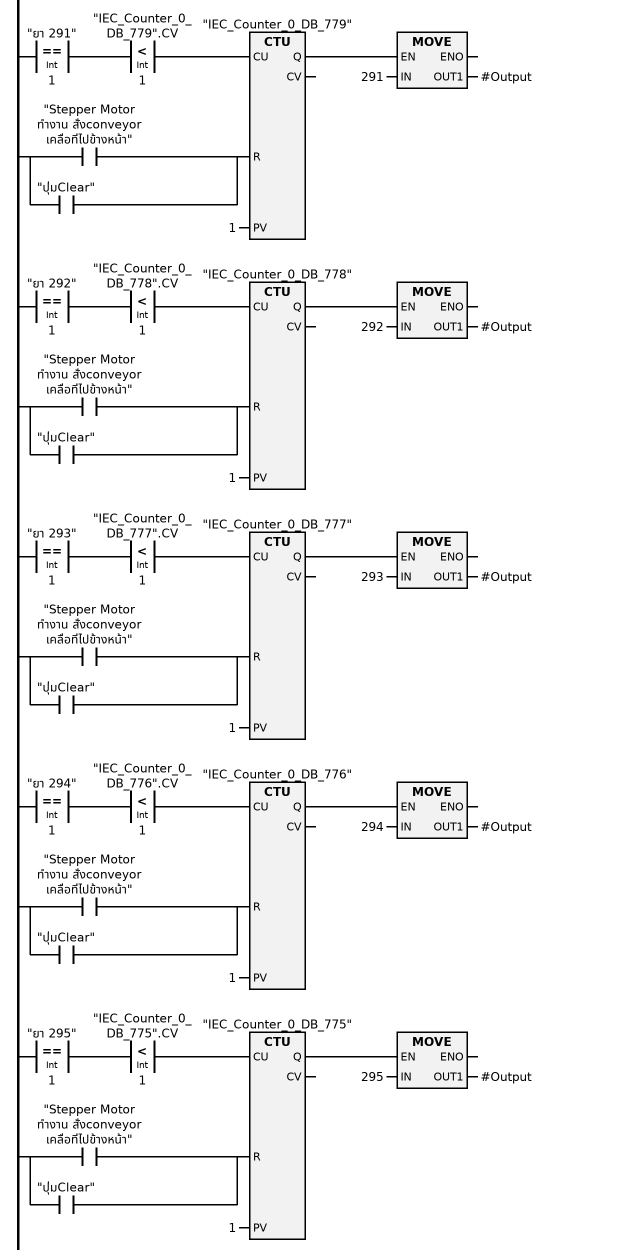
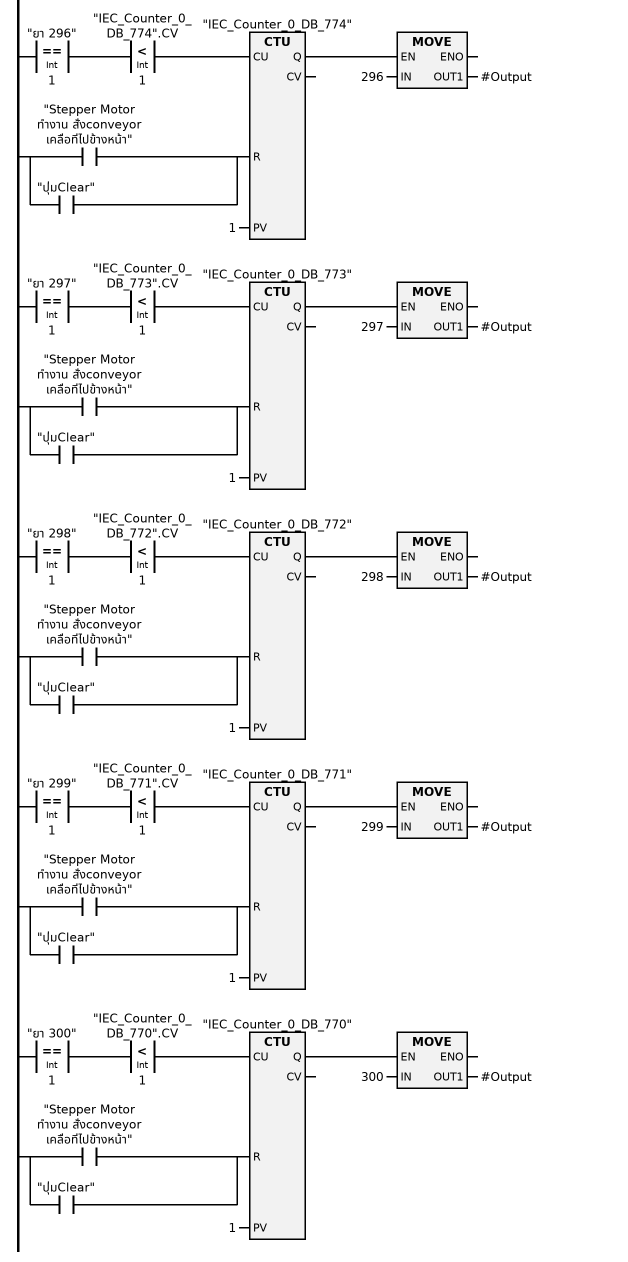
   "IEC_Counter_0_DB_789".CTU(CU := ("ยา 281" = 1) AND ("IEC_Counter_0_DB_789".CV < 1),
                           R := "Stepper Motor ทำงาน สั่งconveyor เคลื่อที่ไปข้างหน้า" OR "ปุ่มClear",
                           PV := 1);
   IF "IEC_Counter_0_DB_789".Q THEN #Output := 281; END_IF;
   "IEC_Counter_0_DB_788".CTU(CU := ("ยา 282" = 1) AND ("IEC_Counter_0_DB_788".CV < 1),
                           R := "Stepper Motor ทำงาน สั่งconveyor เคลื่อที่ไปข้างหน้า" OR "ปุ่มClear",
                           PV := 1);
   IF "IEC_Counter_0_DB_788".Q THEN #Output := 282; END_IF;
   "IEC_Counter_0_DB_787".CTU(CU := ("ยา 283" = 1) AND ("IEC_Counter_0_DB_787".CV < 1),
                           R := "Stepper Motor ทำงาน สั่งconveyor เคลื่อที่ไปข้างหน้า" OR "ปุ่มClear",
                           PV := 1);
   IF "IEC_Counter_0_DB_787".Q THEN #Output := 283; END_IF;
   "IEC_Counter_0_DB_786".CTU(CU := ("ยา 284" = 1) AND ("IEC_Counter_0_DB_786".CV < 1),
                           R := "Stepper Motor ทำงาน สั่งconveyor เคลื่อที่ไปข้างหน้า" OR "ปุ่มClear",
                           PV := 1);
   IF "IEC_Counter_0_DB_786".Q THEN #Output := 284; END_IF;
   "IEC_Counter_0_DB_785".CTU(CU := ("ยา 285" = 1) AND ("IEC_Counter_0_DB_785".CV < 1),
                           R := "Stepper Motor ทำงาน สั่งconveyor เคลื่อที่ไปข้างหน้า" OR "ปุ่มClear",
                           PV := 1);
   IF "IEC_Counter_0_DB_785".Q THEN #Output := 285; END_IF;
   "IEC_Counter_0_DB_784".CTU(CU := ("ยา 286" = 1) AND ("IEC_Counter_0_DB_784".CV < 1),
                           R := "Stepper Motor ทำงาน สั่งconveyor เคลื่อที่ไปข้างหน้า" OR "ปุ่มClear",
                           PV := 1);
   IF "IEC_Counter_0_DB_784".Q THEN #Output := 286; END_IF;
   "IEC_Counter_0_DB_783".CTU(CU := ("ยา 287" = 1) AND ("IEC_Counter_0_DB_783".CV < 1),
                           R := "Stepper Motor ทำงาน สั่งconveyor เคลื่อที่ไปข้างหน้า" OR "ปุ่มClear",
                           PV := 1);
   IF "IEC_Counter_0_DB_783".Q THEN #Output := 287; END_IF;
   "IEC_Counter_0_DB_782".CTU(CU := ("ยา 288" = 1) AND ("IEC_Counter_0_DB_782".CV < 1),
                           R := "Stepper Motor ทำงาน สั่งconveyor เคลื่อที่ไปข้างหน้า" OR "ปุ่มClear",
                           PV := 1);
   IF "IEC_Counter_0_DB_782".Q THEN #Output := 288; END_IF;
   "IEC_Counter_0_DB_781".CTU(CU := ("ยา 289" = 1) AND ("IEC_Counter_0_DB_781".CV < 1),
                           R := "Stepper Motor ทำงาน สั่งconveyor เคลื่อที่ไปข้างหน้า" OR "ปุ่มClear",
                           PV := 1);
   IF "IEC_Counter_0_DB_781".Q THEN #Output := 289; END_IF;
   "IEC_Counter_0_DB_780".CTU(CU := ("ยา 290" = 1) AND ("IEC_Counter_0_DB_780".CV < 1),
                           R := "Stepper Motor ทำงาน สั่งconveyor เคลื่อที่ไปข้างหน้า" OR "ปุ่มClear",
                           PV := 1);
   IF "IEC_Counter_0_DB_780".Q THEN #Output := 290; END_IF;
   "IEC_Counter_0_DB_779".CTU(CU := ("ยา 291" = 1) AND ("IEC_Counter_0_DB_779".CV < 1),
                           R := "Stepper Motor ทำงาน สั่งconveyor เคลื่อที่ไปข้างหน้า" OR "ปุ่มClear",
                           PV := 1);
   IF "IEC_Counter_0_DB_779".Q THEN #Output := 291; END_IF;
   "IEC_Counter_0_DB_778".CTU(CU := ("ยา 292" = 1) AND ("IEC_Counter_0_DB_778".CV < 1),
                           R := "Stepper Motor ทำงาน สั่งconveyor เคลื่อที่ไปข้างหน้า" OR "ปุ่มClear",
                           PV := 1);
   IF "IEC_Counter_0_DB_778".Q THEN #Output := 292; END_IF;
   "IEC_Counter_0_DB_777".CTU(CU := ("ยา 293" = 1) AND ("IEC_Counter_0_DB_777".CV < 1),
                           R := "Stepper Motor ทำงาน สั่งconveyor เคลื่อที่ไปข้างหน้า" OR "ปุ่มClear",
                           PV := 1);
   IF "IEC_Counter_0_DB_777".Q THEN #Output := 293; END_IF;
   "IEC_Counter_0_DB_776".CTU(CU := ("ยา 294" = 1) AND ("IEC_Counter_0_DB_776".CV < 1),
                           R := "Stepper Motor ทำงาน สั่งconveyor เคลื่อที่ไปข้างหน้า" OR "ปุ่มClear",
                           PV := 1);
   IF "IEC_Counter_0_DB_776".Q THEN #Output := 294; END_IF;
   "IEC_Counter_0_DB_775".CTU(CU := ("ยา 295" = 1) AND ("IEC_Counter_0_DB_775".CV < 1),
                           R := "Stepper Motor ทำงาน สั่งconveyor เคลื่อที่ไปข้างหน้า" OR "ปุ่มClear",
                           PV := 1);
   IF "IEC_Counter_0_DB_775".Q THEN #Output := 295; END_IF;
   "IEC_Counter_0_DB_774".CTU(CU := ("ยา 296" = 1) AND ("IEC_Counter_0_DB_774".CV < 1),
                           R := "Stepper Motor ทำงาน สั่งconveyor เคลื่อที่ไปข้างหน้า" OR "ปุ่มClear",
                           PV := 1);
   IF "IEC_Counter_0_DB_774".Q THEN #Output := 296; END_IF;
   "IEC_Counter_0_DB_773".CTU(CU := ("ยา 297" = 1) AND ("IEC_Counter_0_DB_773".CV < 1),
                           R := "Stepper Motor ทำงาน สั่งconveyor เคลื่อที่ไปข้างหน้า" OR "ปุ่มClear",
                           PV := 1);
   IF "IEC_Counter_0_DB_773".Q THEN #Output := 297; END_IF;
   "IEC_Counter_0_DB_772".CTU(CU := ("ยา 298" = 1) AND ("IEC_Counter_0_DB_772".CV < 1),
                           R := "Stepper Motor ทำงาน สั่งconveyor เคลื่อที่ไปข้างหน้า" OR "ปุ่มClear",
                           PV := 1);
   IF "IEC_Counter_0_DB_772".Q THEN #Output := 298; END_IF;
   "IEC_Counter_0_DB_771".CTU(CU := ("ยา 299" = 1) AND ("IEC_Counter_0_DB_771".CV < 1),
                           R := "Stepper Motor ทำงาน สั่งconveyor เคลื่อที่ไปข้างหน้า" OR "ปุ่มClear",
                           PV := 1);
   IF "IEC_Counter_0_DB_771".Q THEN #Output := 299; END_IF;
   "IEC_Counter_0_DB_770".CTU(CU := ("ยา 300" = 1) AND ("IEC_Counter_0_DB_770".CV < 1),
                           R := "Stepper Motor ทำงาน สั่งconveyor เคลื่อที่ไปข้างหน้า" OR "ปุ่มClear",
                           PV := 1);
   IF "IEC_Counter_0_DB_770".Q THEN #Output := 300; END_IF;
END_REGION

REGION Network 16
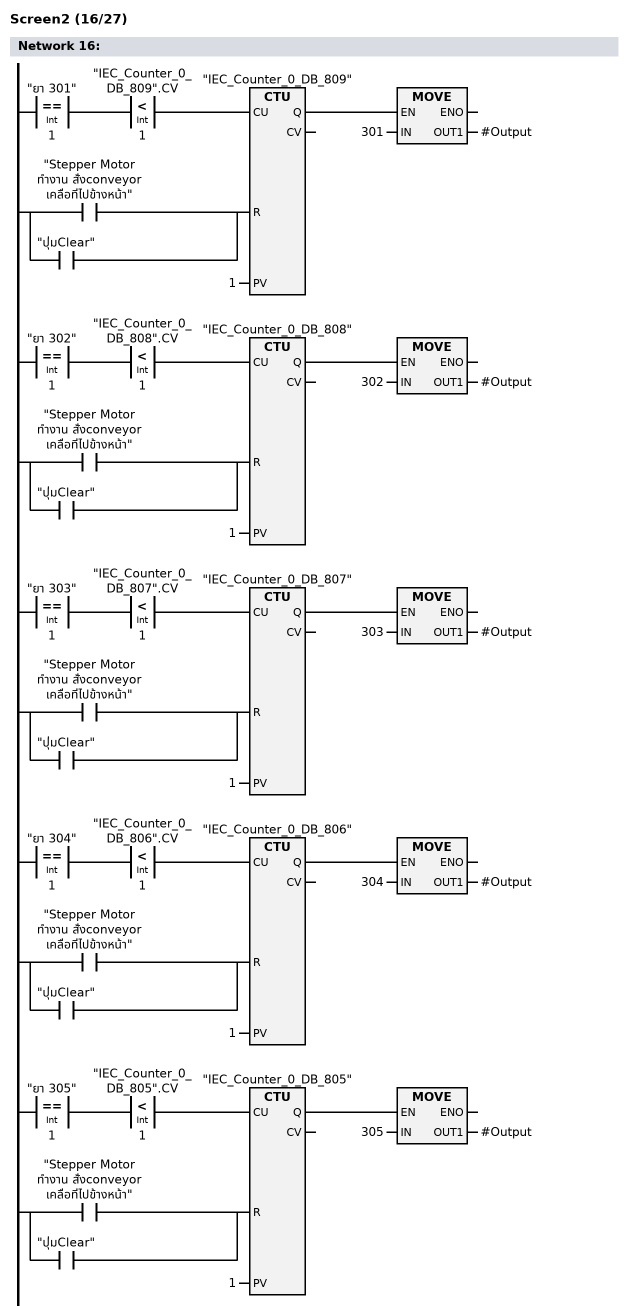
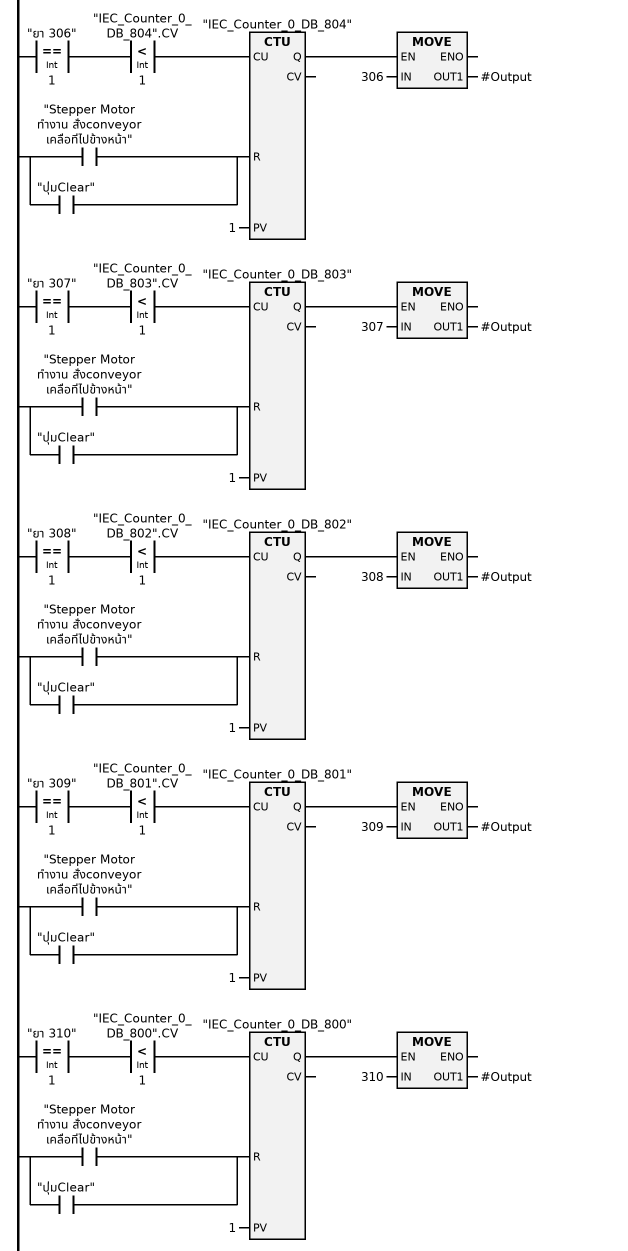
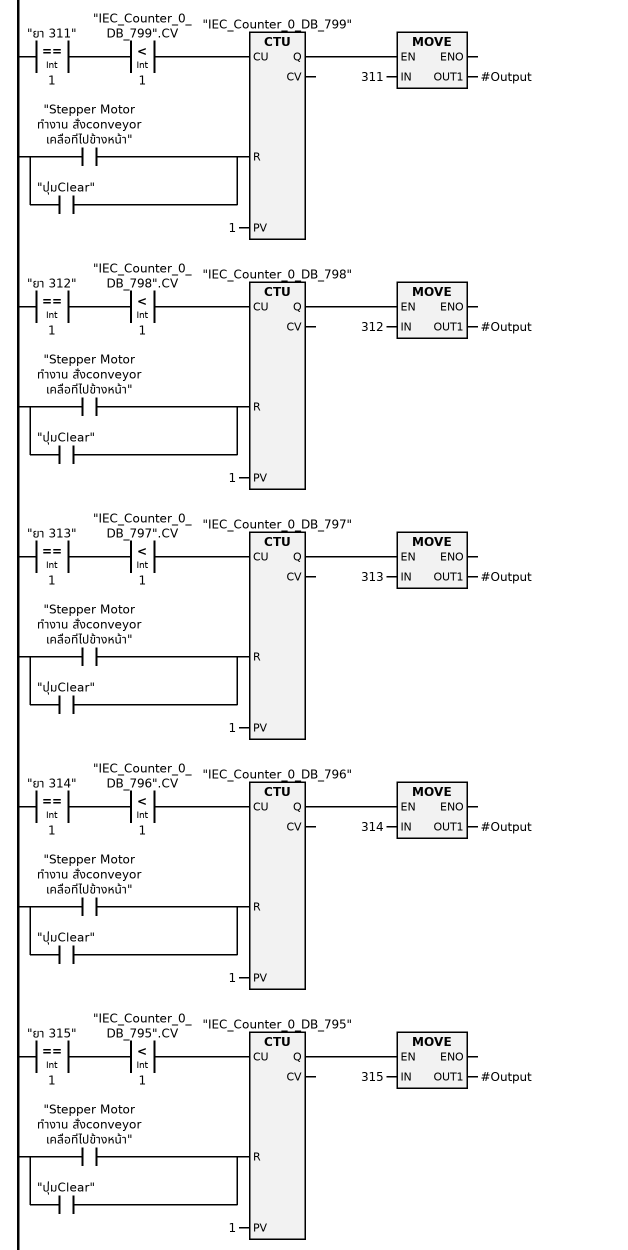
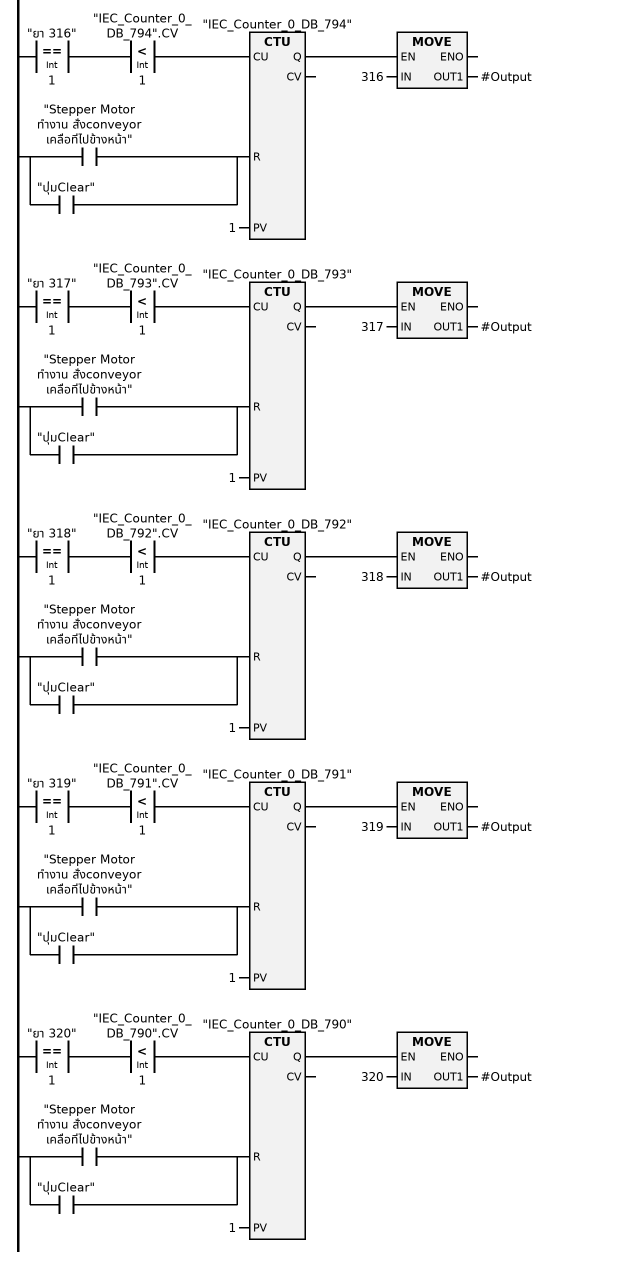
   "IEC_Counter_0_DB_809".CTU(CU := ("ยา 301" = 1) AND ("IEC_Counter_0_DB_809".CV < 1),
                           R := "Stepper Motor ทำงาน สั่งconveyor เคลื่อที่ไปข้างหน้า" OR "ปุ่มClear",
                           PV := 1);
   IF "IEC_Counter_0_DB_809".Q THEN #Output := 301; END_IF;
   "IEC_Counter_0_DB_808".CTU(CU := ("ยา 302" = 1) AND ("IEC_Counter_0_DB_808".CV < 1),
                           R := "Stepper Motor ทำงาน สั่งconveyor เคลื่อที่ไปข้างหน้า" OR "ปุ่มClear",
                           PV := 1);
   IF "IEC_Counter_0_DB_808".Q THEN #Output := 302; END_IF;
   "IEC_Counter_0_DB_807".CTU(CU := ("ยา 303" = 1) AND ("IEC_Counter_0_DB_807".CV < 1),
                           R := "Stepper Motor ทำงาน สั่งconveyor เคลื่อที่ไปข้างหน้า" OR "ปุ่มClear",
                           PV := 1);
   IF "IEC_Counter_0_DB_807".Q THEN #Output := 303; END_IF;
   "IEC_Counter_0_DB_806".CTU(CU := ("ยา 304" = 1) AND ("IEC_Counter_0_DB_806".CV < 1),
                           R := "Stepper Motor ทำงาน สั่งconveyor เคลื่อที่ไปข้างหน้า" OR "ปุ่มClear",
                           PV := 1);
   IF "IEC_Counter_0_DB_806".Q THEN #Output := 304; END_IF;
   "IEC_Counter_0_DB_805".CTU(CU := ("ยา 305" = 1) AND ("IEC_Counter_0_DB_805".CV < 1),
                           R := "Stepper Motor ทำงาน สั่งconveyor เคลื่อที่ไปข้างหน้า" OR "ปุ่มClear",
                           PV := 1);
   IF "IEC_Counter_0_DB_805".Q THEN #Output := 305; END_IF;
   "IEC_Counter_0_DB_804".CTU(CU := ("ยา 306" = 1) AND ("IEC_Counter_0_DB_804".CV < 1),
                           R := "Stepper Motor ทำงาน สั่งconveyor เคลื่อที่ไปข้างหน้า" OR "ปุ่มClear",
                           PV := 1);
   IF "IEC_Counter_0_DB_804".Q THEN #Output := 306; END_IF;
   "IEC_Counter_0_DB_803".CTU(CU := ("ยา 307" = 1) AND ("IEC_Counter_0_DB_803".CV < 1),
                           R := "Stepper Motor ทำงาน สั่งconveyor เคลื่อที่ไปข้างหน้า" OR "ปุ่มClear",
                           PV := 1);
   IF "IEC_Counter_0_DB_803".Q THEN #Output := 307; END_IF;
   "IEC_Counter_0_DB_802".CTU(CU := ("ยา 308" = 1) AND ("IEC_Counter_0_DB_802".CV < 1),
                           R := "Stepper Motor ทำงาน สั่งconveyor เคลื่อที่ไปข้างหน้า" OR "ปุ่มClear",
                           PV := 1);
   IF "IEC_Counter_0_DB_802".Q THEN #Output := 308; END_IF;
   "IEC_Counter_0_DB_801".CTU(CU := ("ยา 309" = 1) AND ("IEC_Counter_0_DB_801".CV < 1),
                           R := "Stepper Motor ทำงาน สั่งconveyor เคลื่อที่ไปข้างหน้า" OR "ปุ่มClear",
                           PV := 1);
   IF "IEC_Counter_0_DB_801".Q THEN #Output := 309; END_IF;
   "IEC_Counter_0_DB_800".CTU(CU := ("ยา 310" = 1) AND ("IEC_Counter_0_DB_800".CV < 1),
                           R := "Stepper Motor ทำงาน สั่งconveyor เคลื่อที่ไปข้างหน้า" OR "ปุ่มClear",
                           PV := 1);
   IF "IEC_Counter_0_DB_800".Q THEN #Output := 310; END_IF;
   "IEC_Counter_0_DB_799".CTU(CU := ("ยา 311" = 1) AND ("IEC_Counter_0_DB_799".CV < 1),
                           R := "Stepper Motor ทำงาน สั่งconveyor เคลื่อที่ไปข้างหน้า" OR "ปุ่มClear",
                           PV := 1);
   IF "IEC_Counter_0_DB_799".Q THEN #Output := 311; END_IF;
   "IEC_Counter_0_DB_798".CTU(CU := ("ยา 312" = 1) AND ("IEC_Counter_0_DB_798".CV < 1),
                           R := "Stepper Motor ทำงาน สั่งconveyor เคลื่อที่ไปข้างหน้า" OR "ปุ่มClear",
                           PV := 1);
   IF "IEC_Counter_0_DB_798".Q THEN #Output := 312; END_IF;
   "IEC_Counter_0_DB_797".CTU(CU := ("ยา 313" = 1) AND ("IEC_Counter_0_DB_797".CV < 1),
                           R := "Stepper Motor ทำงาน สั่งconveyor เคลื่อที่ไปข้างหน้า" OR "ปุ่มClear",
                           PV := 1);
   IF "IEC_Counter_0_DB_797".Q THEN #Output := 313; END_IF;
   "IEC_Counter_0_DB_796".CTU(CU := ("ยา 314" = 1) AND ("IEC_Counter_0_DB_796".CV < 1),
                           R := "Stepper Motor ทำงาน สั่งconveyor เคลื่อที่ไปข้างหน้า" OR "ปุ่มClear",
                           PV := 1);
   IF "IEC_Counter_0_DB_796".Q THEN #Output := 314; END_IF;
   "IEC_Counter_0_DB_795".CTU(CU := ("ยา 315" = 1) AND ("IEC_Counter_0_DB_795".CV < 1),
                           R := "Stepper Motor ทำงาน สั่งconveyor เคลื่อที่ไปข้างหน้า" OR "ปุ่มClear",
                           PV := 1);
   IF "IEC_Counter_0_DB_795".Q THEN #Output := 315; END_IF;
   "IEC_Counter_0_DB_794".CTU(CU := ("ยา 316" = 1) AND ("IEC_Counter_0_DB_794".CV < 1),
                           R := "Stepper Motor ทำงาน สั่งconveyor เคลื่อที่ไปข้างหน้า" OR "ปุ่มClear",
                           PV := 1);
   IF "IEC_Counter_0_DB_794".Q THEN #Output := 316; END_IF;
   "IEC_Counter_0_DB_793".CTU(CU := ("ยา 317" = 1) AND ("IEC_Counter_0_DB_793".CV < 1),
                           R := "Stepper Motor ทำงาน สั่งconveyor เคลื่อที่ไปข้างหน้า" OR "ปุ่มClear",
                           PV := 1);
   IF "IEC_Counter_0_DB_793".Q THEN #Output := 317; END_IF;
   "IEC_Counter_0_DB_792".CTU(CU := ("ยา 318" = 1) AND ("IEC_Counter_0_DB_792".CV < 1),
                           R := "Stepper Motor ทำงาน สั่งconveyor เคลื่อที่ไปข้างหน้า" OR "ปุ่มClear",
                           PV := 1);
   IF "IEC_Counter_0_DB_792".Q THEN #Output := 318; END_IF;
   "IEC_Counter_0_DB_791".CTU(CU := ("ยา 319" = 1) AND ("IEC_Counter_0_DB_791".CV < 1),
                           R := "Stepper Motor ทำงาน สั่งconveyor เคลื่อที่ไปข้างหน้า" OR "ปุ่มClear",
                           PV := 1);
   IF "IEC_Counter_0_DB_791".Q THEN #Output := 319; END_IF;
   "IEC_Counter_0_DB_790".CTU(CU := ("ยา 320" = 1) AND ("IEC_Counter_0_DB_790".CV < 1),
                           R := "Stepper Motor ทำงาน สั่งconveyor เคลื่อที่ไปข้างหน้า" OR "ปุ่มClear",
                           PV := 1);
   IF "IEC_Counter_0_DB_790".Q THEN #Output := 320; END_IF;
END_REGION

REGION Network 17
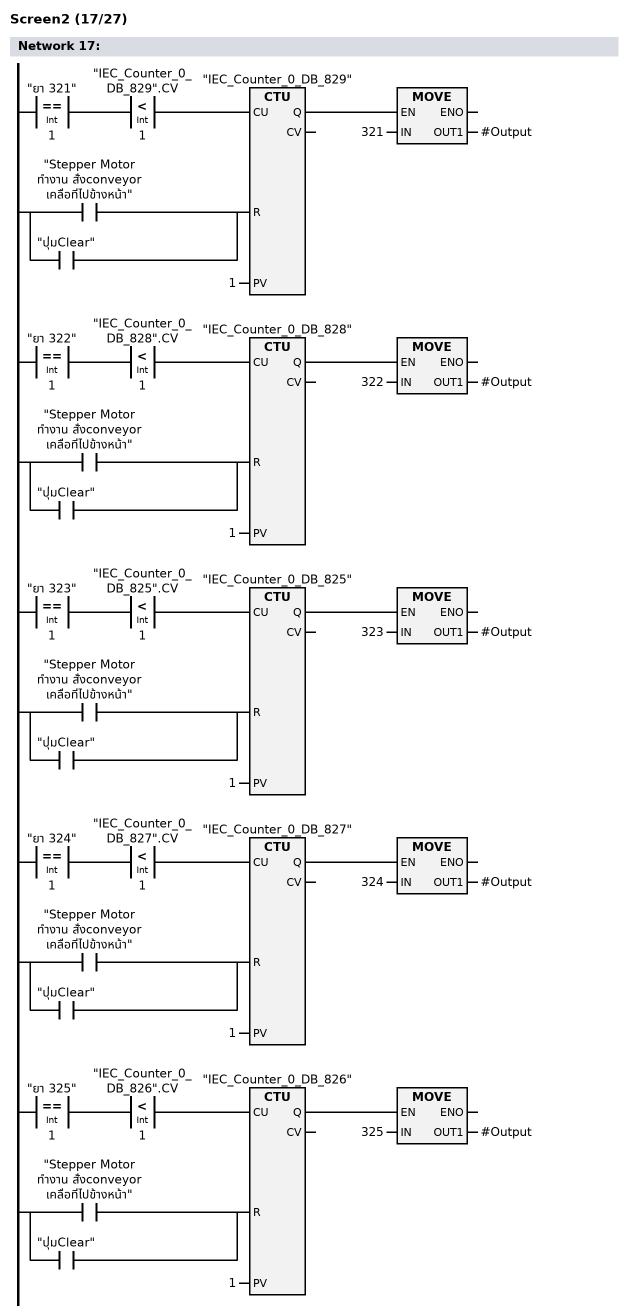
